//     PlcTask Inputs/GVL_iXlinker.Device_2_EtherCAT.Term_9_EK1100.Term_34_EL3403.PM_Inputs_Channel_1.TxPDO_Toggle <-> PM Inputs Channel 1/TxPDO Toggle
//     PlcTask Inputs/GVL_iXlinker.Device_2_EtherCAT.Term_9_EK1100.Term_34_EL3403.PM_Inputs_Channel_2.TxPDO_Toggle <-> PM Inputs Channel 2/TxPDO Toggle
//     PlcTask Inputs/GVL_iXlinker.Device_2_EtherCAT.Term_9_EK1100.Term_34_EL3403.PM_Inputs_Channel_3.TxPDO_Toggle <-> PM Inputs Channel 3/TxPDO Toggle
//     PlcTask Inputs/GVL_iXlinker.Device_2_EtherCAT.Term_9_EK1100.Term_34_EL3403.PM_Inputs_Channel_1.Variant_value <-> PM Inputs Channel 1/Variant value
//     PlcTask Inputs/GVL_iXlinker.Device_2_EtherCAT.Term_9_EK1100.Term_34_EL3403.PM_Inputs_Channel_2.Variant_value <-> PM Inputs Channel 2/Variant value
//     PlcTask Inputs/GVL_iXlinker.Device_2_EtherCAT.Term_9_EK1100.Term_34_EL3403.PM_Inputs_Channel_3.Variant_value <-> PM Inputs Channel 3/Variant value
//     PlcTask Inputs/GVL_iXlinker.Device_2_EtherCAT.Term_9_EK1100.Term_34_EL3403.PM_Inputs_Channel_1.Voltage <-> PM Inputs Channel 1/Voltage
//     PlcTask Inputs/GVL_iXlinker.Device_2_EtherCAT.Term_9_EK1100.Term_34_EL3403.PM_Inputs_Channel_2.Voltage <-> PM Inputs Channel 2/Voltage
//     PlcTask Inputs/GVL_iXlinker.Device_2_EtherCAT.Term_9_EK1100.Term_34_EL3403.PM_Inputs_Channel_3.Voltage <-> PM Inputs Channel 3/Voltage
//     PlcTask Inputs/GVL_iXlinker.Device_2_EtherCAT.Term_9_EK1100.Term_34_EL3403.PM_Status_data.Missing_zero_crossing_A <-> PM Status data/Missing zero crossing A
//     PlcTask Inputs/GVL_iXlinker.Device_2_EtherCAT.Term_9_EK1100.Term_34_EL3403.PM_Status_data.Missing_zero_crossing_B <-> PM Status data/Missing zero crossing B
//     PlcTask Inputs/GVL_iXlinker.Device_2_EtherCAT.Term_9_EK1100.Term_34_EL3403.PM_Status_data.Missing_zero_crossing_C <-> PM Status data/Missing zero crossing C
//     PlcTask Inputs/GVL_iXlinker.Device_2_EtherCAT.Term_9_EK1100.Term_34_EL3403.PM_Status_data.Phase_sequence_error <-> PM Status data/Phase sequence error
//     PlcTask Inputs/GVL_iXlinker.Device_2_EtherCAT.Term_9_EK1100.Term_34_EL3403.WcState.InputToggle <-> WcState/InputToggle
//     PlcTask Inputs/GVL_iXlinker.Device_2_EtherCAT.Term_9_EK1100.Term_34_EL3403.WcState.WcState <-> WcState/WcState
//     PlcTask Outputs/GVL_iXlinker.Device_2_EtherCAT.Term_9_EK1100.Term_34_EL3403.PM_Outputs_Channel_1.Index <-> PM Outputs Channel 1/Index
//     PlcTask Outputs/GVL_iXlinker.Device_2_EtherCAT.Term_9_EK1100.Term_34_EL3403.PM_Outputs_Channel_2.Index <-> PM Outputs Channel 2/Index
//     PlcTask Outputs/GVL_iXlinker.Device_2_EtherCAT.Term_9_EK1100.Term_34_EL3403.PM_Outputs_Channel_3.Index <-> PM Outputs Channel 3/Index
//   TcoIoTests/TcoIoTests Instance <-> Device 2 (EtherCAT)/Term 9 (EK1100)/Term 35 (EL6001)
//     PlcTask Inputs/GVL_iXlinker.Device_2_EtherCAT.Term_9_EK1100.Term_35_EL6001.COM_Inputs.Data_In[{0..21}] <-> COM Inputs/Data In {0..21}  (22 links)
//     PlcTask Inputs/GVL_iXlinker.Device_2_EtherCAT.Term_9_EK1100.Term_35_EL6001.COM_Inputs.Status/Buffer_full <-> COM Inputs/Status/Buffer full
//     PlcTask Inputs/GVL_iXlinker.Device_2_EtherCAT.Term_9_EK1100.Term_35_EL6001.COM_Inputs.Status/Framing_error <-> COM Inputs/Status/Framing error
//     PlcTask Inputs/GVL_iXlinker.Device_2_EtherCAT.Term_9_EK1100.Term_35_EL6001.COM_Inputs.Status/Init_accepted <-> COM Inputs/Status/Init accepted
//     PlcTask Inputs/GVL_iXlinker.Device_2_EtherCAT.Term_9_EK1100.Term_35_EL6001.COM_Inputs.Status/Input_length <-> COM Inputs/Status/Input length
//     PlcTask Inputs/GVL_iXlinker.Device_2_EtherCAT.Term_9_EK1100.Term_35_EL6001.COM_Inputs.Status/Overrun_error <-> COM Inputs/Status/Overrun error
//     PlcTask Inputs/GVL_iXlinker.Device_2_EtherCAT.Term_9_EK1100.Term_35_EL6001.COM_Inputs.Status/Parity_error <-> COM Inputs/Status/Parity error
//     PlcTask Inputs/GVL_iXlinker.Device_2_EtherCAT.Term_9_EK1100.Term_35_EL6001.COM_Inputs.Status/Receive_request <-> COM Inputs/Status/Receive request
//     PlcTask Inputs/GVL_iXlinker.Device_2_EtherCAT.Term_9_EK1100.Term_35_EL6001.COM_Inputs.Status/Transmit_accepted <-> COM Inputs/Status/Transmit accepted
//     PlcTask Inputs/GVL_iXlinker.Device_2_EtherCAT.Term_9_EK1100.Term_35_EL6001.InfoData.AdsAddr <-> InfoData/AdsAddr
//     PlcTask Inputs/GVL_iXlinker.Device_2_EtherCAT.Term_9_EK1100.Term_35_EL6001.InfoData.State <-> InfoData/State
//     PlcTask Inputs/GVL_iXlinker.Device_2_EtherCAT.Term_9_EK1100.Term_35_EL6001.WcState.InputToggle <-> WcState/InputToggle
//     PlcTask Inputs/GVL_iXlinker.Device_2_EtherCAT.Term_9_EK1100.Term_35_EL6001.WcState.WcState <-> WcState/WcState
//     PlcTask Outputs/GVL_iXlinker.Device_2_EtherCAT.Term_9_EK1100.Term_35_EL6001.COM_Outputs.Ctrl/Init_request <-> COM Outputs/Ctrl/Init request
//     PlcTask Outputs/GVL_iXlinker.Device_2_EtherCAT.Term_9_EK1100.Term_35_EL6001.COM_Outputs.Ctrl/Output_length <-> COM Outputs/Ctrl/Output length
//     PlcTask Outputs/GVL_iXlinker.Device_2_EtherCAT.Term_9_EK1100.Term_35_EL6001.COM_Outputs.Ctrl/Receive_accepted <-> COM Outputs/Ctrl/Receive accepted
//     PlcTask Outputs/GVL_iXlinker.Device_2_EtherCAT.Term_9_EK1100.Term_35_EL6001.COM_Outputs.Ctrl/Send_continues <-> COM Outputs/Ctrl/Send continues
//     PlcTask Outputs/GVL_iXlinker.Device_2_EtherCAT.Term_9_EK1100.Term_35_EL6001.COM_Outputs.Ctrl/Transmit_request <-> COM Outputs/Ctrl/Transmit request
//     PlcTask Outputs/GVL_iXlinker.Device_2_EtherCAT.Term_9_EK1100.Term_35_EL6001.COM_Outputs.Data_Out[{0..21}] <-> COM Outputs/Data Out {0..21}  (22 links)
//   TcoIoTests/TcoIoTests Instance <-> Device 2 (EtherCAT)/Term 9 (EK1100)/Term 36 (EL3024)
//     PlcTask Inputs/GVL_iXlinker.Device_2_EtherCAT.Term_9_EK1100.Term_36_EL3024.AI_Standard_Channel_{1..4}.Status/Error <-> AI Standard Channel {1..4}/Status/Error  (4 links)
//     PlcTask Inputs/GVL_iXlinker.Device_2_EtherCAT.Term_9_EK1100.Term_36_EL3024.AI_Standard_Channel_1.Status/Limit_1 <-> AI Standard Channel 1/Status/Limit 1
//     PlcTask Inputs/GVL_iXlinker.Device_2_EtherCAT.Term_9_EK1100.Term_36_EL3024.AI_Standard_Channel_1.Status/Limit_2 <-> AI Standard Channel 1/Status/Limit 2
//     PlcTask Inputs/GVL_iXlinker.Device_2_EtherCAT.Term_9_EK1100.Term_36_EL3024.AI_Standard_Channel_2.Status/Limit_1 <-> AI Standard Channel 2/Status/Limit 1
//     PlcTask Inputs/GVL_iXlinker.Device_2_EtherCAT.Term_9_EK1100.Term_36_EL3024.AI_Standard_Channel_2.Status/Limit_2 <-> AI Standard Channel 2/Status/Limit 2
//     PlcTask Inputs/GVL_iXlinker.Device_2_EtherCAT.Term_9_EK1100.Term_36_EL3024.AI_Standard_Channel_3.Status/Limit_1 <-> AI Standard Channel 3/Status/Limit 1
//     PlcTask Inputs/GVL_iXlinker.Device_2_EtherCAT.Term_9_EK1100.Term_36_EL3024.AI_Standard_Channel_3.Status/Limit_2 <-> AI Standard Channel 3/Status/Limit 2
//     PlcTask Inputs/GVL_iXlinker.Device_2_EtherCAT.Term_9_EK1100.Term_36_EL3024.AI_Standard_Channel_4.Status/Limit_1 <-> AI Standard Channel 4/Status/Limit 1
//     PlcTask Inputs/GVL_iXlinker.Device_2_EtherCAT.Term_9_EK1100.Term_36_EL3024.AI_Standard_Channel_4.Status/Limit_2 <-> AI Standard Channel 4/Status/Limit 2
//     PlcTask Inputs/GVL_iXlinker.Device_2_EtherCAT.Term_9_EK1100.Term_36_EL3024.AI_Standard_Channel_{1..4}.Status/Overrange <-> AI Standard Channel {1..4}/Status/Overrange  (4 links)
//     PlcTask Inputs/GVL_iXlinker.Device_2_EtherCAT.Term_9_EK1100.Term_36_EL3024.AI_Standard_Channel_{1..4}.Status/TxPDO_State <-> AI Standard Channel {1..4}/Status/TxPDO State  (4 links)
//     PlcTask Inputs/GVL_iXlinker.Device_2_EtherCAT.Term_9_EK1100.Term_36_EL3024.AI_Standard_Channel_{1..4}.Status/TxPDO_Toggle <-> AI Standard Channel {1..4}/Status/TxPDO Toggle  (4 links)
//     PlcTask Inputs/GVL_iXlinker.Device_2_EtherCAT.Term_9_EK1100.Term_36_EL3024.AI_Standard_Channel_{1..4}.Status/Underrange <-> AI Standard Channel {1..4}/Status/Underrange  (4 links)
//     PlcTask Inputs/GVL_iXlinker.Device_2_EtherCAT.Term_9_EK1100.Term_36_EL3024.AI_Standard_Channel_{1..4}.Value <-> AI Standard Channel {1..4}/Value  (4 links)
//     PlcTask Inputs/GVL_iXlinker.Device_2_EtherCAT.Term_9_EK1100.Term_36_EL3024.InfoData.AdsAddr <-> InfoData/AdsAddr
//     PlcTask Inputs/GVL_iXlinker.Device_2_EtherCAT.Term_9_EK1100.Term_36_EL3024.InfoData.State <-> InfoData/State
//     PlcTask Inputs/GVL_iXlinker.Device_2_EtherCAT.Term_9_EK1100.Term_36_EL3024.WcState.InputToggle <-> WcState/InputToggle
//     PlcTask Inputs/GVL_iXlinker.Device_2_EtherCAT.Term_9_EK1100.Term_36_EL3024.WcState.WcState <-> WcState/WcState
//   TcoIoTests/TcoIoTests Instance <-> Device 3 (EtherCAT)
//     PlcTask Inputs/GVL_iXlinker.Device_3_EtherCAT.InfoData.AmsNetId <-> InfoData/AmsNetId
//     PlcTask Inputs/GVL_iXlinker.Device_3_EtherCAT.InfoData.CfgSlaveCount <-> InfoData/CfgSlaveCount
//     PlcTask Inputs/GVL_iXlinker.Device_3_EtherCAT.InfoData.ChangeCount <-> InfoData/ChangeCount
//     PlcTask Inputs/GVL_iXlinker.Device_3_EtherCAT.InfoData.DevId <-> InfoData/DevId
//     PlcTask Inputs/GVL_iXlinker.Device_3_EtherCAT.Inputs.DevState <-> Inputs/DevState
//     PlcTask Inputs/GVL_iXlinker.Device_3_EtherCAT.Inputs.Frm0InputToggle <-> Inputs/Frm0InputToggle
//     PlcTask Inputs/GVL_iXlinker.Device_3_EtherCAT.Inputs.Frm0State <-> Inputs/Frm0State
//     PlcTask Inputs/GVL_iXlinker.Device_3_EtherCAT.Inputs.Frm0WcState <-> Inputs/Frm0WcState
//     PlcTask Inputs/GVL_iXlinker.Device_3_EtherCAT.Inputs.SlaveCount <-> Inputs/SlaveCount
//     PlcTask Outputs/GVL_iXlinker.Device_3_EtherCAT.Outputs.DevCtrl <-> Outputs/DevCtrl
//     PlcTask Outputs/GVL_iXlinker.Device_3_EtherCAT.Outputs.Frm0Ctrl <-> Outputs/Frm0Ctrl
//     PlcTask Outputs/GVL_iXlinker.Device_3_EtherCAT.Outputs.Frm0WcCtrl <-> Outputs/Frm0WcCtrl
//   TcoIoTests/TcoIoTests Instance <-> Device 3 (EtherCAT)/Term 146 (EK1100)
//     PlcTask Inputs/GVL_iXlinker.Device_3_EtherCAT.Term_146_EK1100.InfoData.State <-> InfoData/State
//   TcoIoTests/TcoIoTests Instance <-> Device 3 (EtherCAT)/Term 146 (EK1100)/Term 147 (EK1122)
//     PlcTask Inputs/GVL_iXlinker.Device_3_EtherCAT.Term_146_EK1100.Term_147_EK1122.InfoData.State <-> InfoData/State
//   TcoIoTests/TcoIoTests Instance <-> Device 3 (EtherCAT)/Term 146 (EK1100)/Term 147 (EK1122)/Term 153 (EK1100)
//     PlcTask Inputs/GVL_iXlinker.Device_3_EtherCAT.Term_146_EK1100.Term_147_EK1122.Term_153_EK1100.InfoData.State <-> InfoData/State
//   TcoIoTests/TcoIoTests Instance <-> Device 3 (EtherCAT)/Term 146 (EK1100)/Term 147 (EK1122)/Term 153 (EK1100)/Term 154 (EK1122)
//     PlcTask Inputs/GVL_iXlinker.Device_3_EtherCAT.Term_146_EK1100.Term_147_EK1122.Term_153_EK1100.Term_154_EK1122.InfoData.State <-> InfoData/State
//   TcoIoTests/TcoIoTests Instance <-> Device 3 (EtherCAT)/Term 146 (EK1100)/Term 147 (EK1122)/Term 153 (EK1100)/Term 154 (EK1122)/Term 157 (EK1100)
//     PlcTask Inputs/GVL_iXlinker.Device_3_EtherCAT.Term_146_EK1100.Term_147_EK1122.Term_153_EK1100.Term_154_EK1122.Term_157_EK1100.InfoData.State <-> InfoData/State
//   TcoIoTests/TcoIoTests Instance <-> Device 3 (EtherCAT)/Term 146 (EK1100)/Term 147 (EK1122)/Term 153 (EK1100)/Term 154 (EK1122)/Term 157 (EK1100)/Term 159 (EL1809)
//     PlcTask Inputs/GVL_iXlinker.Device_3_EtherCAT.Term_146_EK1100.Term_147_EK1122.Term_153_EK1100.Term_154_EK1122.Term_157_EK1100.Term_159_EL1809.Channel_{1..16}.Input <-> Channel {1..16}/Input  (16 links)
//     PlcTask Inputs/GVL_iXlinker.Device_3_EtherCAT.Term_146_EK1100.Term_147_EK1122.Term_153_EK1100.Term_154_EK1122.Term_157_EK1100.Term_159_EL1809.InfoData.State <-> InfoData/State
//     PlcTask Inputs/GVL_iXlinker.Device_3_EtherCAT.Term_146_EK1100.Term_147_EK1122.Term_153_EK1100.Term_154_EK1122.Term_157_EK1100.Term_159_EL1809.WcState.InputToggle <-> WcState/InputToggle
//     PlcTask Inputs/GVL_iXlinker.Device_3_EtherCAT.Term_146_EK1100.Term_147_EK1122.Term_153_EK1100.Term_154_EK1122.Term_157_EK1100.Term_159_EL1809.WcState.WcState <-> WcState/WcState
//   TcoIoTests/TcoIoTests Instance <-> Device 3 (EtherCAT)/Term 146 (EK1100)/Term 147 (EK1122)/Term 153 (EK1100)/Term 154 (EK1122)/Term 158 (EK1100)
//     PlcTask Inputs/GVL_iXlinker.Device_3_EtherCAT.Term_146_EK1100.Term_147_EK1122.Term_153_EK1100.Term_154_EK1122.Term_158_EK1100.InfoData.State <-> InfoData/State
//   TcoIoTests/TcoIoTests Instance <-> Device 3 (EtherCAT)/Term 146 (EK1100)/Term 147 (EK1122)/Term 153 (EK1100)/Term 154 (EK1122)/Term 158 (EK1100)/Term 160 (EL1809)
//     PlcTask Inputs/GVL_iXlinker.Device_3_EtherCAT.Term_146_EK1100.Term_147_EK1122.Term_153_EK1100.Term_154_EK1122.Term_158_EK1100.Term_160_EL1809.Channel_{1..16}.Input <-> Channel {1..16}/Input  (16 links)
//     PlcTask Inputs/GVL_iXlinker.Device_3_EtherCAT.Term_146_EK1100.Term_147_EK1122.Term_153_EK1100.Term_154_EK1122.Term_158_EK1100.Term_160_EL1809.InfoData.State <-> InfoData/State
//     PlcTask Inputs/GVL_iXlinker.Device_3_EtherCAT.Term_146_EK1100.Term_147_EK1122.Term_153_EK1100.Term_154_EK1122.Term_158_EK1100.Term_160_EL1809.WcState.InputToggle <-> WcState/InputToggle
//     PlcTask Inputs/GVL_iXlinker.Device_3_EtherCAT.Term_146_EK1100.Term_147_EK1122.Term_153_EK1100.Term_154_EK1122.Term_158_EK1100.Term_160_EL1809.WcState.WcState <-> WcState/WcState
//   TcoIoTests/TcoIoTests Instance <-> Device 3 (EtherCAT)/Term 146 (EK1100)/Term 147 (EK1122)/Term 153 (EK1100)/Term 155 (EL2008)
//     PlcTask Inputs/GVL_iXlinker.Device_3_EtherCAT.Term_146_EK1100.Term_147_EK1122.Term_153_EK1100.Term_155_EL2008.InfoData.State <-> InfoData/State
//     PlcTask Inputs/GVL_iXlinker.Device_3_EtherCAT.Term_146_EK1100.Term_147_EK1122.Term_153_EK1100.Term_155_EL2008.WcState.WcState <-> WcState/WcState
//     PlcTask Outputs/GVL_iXlinker.Device_3_EtherCAT.Term_146_EK1100.Term_147_EK1122.Term_153_EK1100.Term_155_EL2008.Channel_{1..8}.Output <-> Channel {1..8}/Output  (8 links)
//   TcoIoTests/TcoIoTests Instance <-> Device 3 (EtherCAT)/Term 146 (EK1100)/Term 147 (EK1122)/Term 153 (EK1100)/Term 156 (EL2008)
//     PlcTask Inputs/GVL_iXlinker.Device_3_EtherCAT.Term_146_EK1100.Term_147_EK1122.Term_153_EK1100.Term_156_EL2008.InfoData.State <-> InfoData/State
//     PlcTask Inputs/GVL_iXlinker.Device_3_EtherCAT.Term_146_EK1100.Term_147_EK1122.Term_153_EK1100.Term_156_EL2008.WcState.WcState <-> WcState/WcState
//     PlcTask Outputs/GVL_iXlinker.Device_3_EtherCAT.Term_146_EK1100.Term_147_EK1122.Term_153_EK1100.Term_156_EL2008.Channel_{1..8}.Output <-> Channel {1..8}/Output  (8 links)
//   TcoIoTests/TcoIoTests Instance <-> Device 3 (EtherCAT)/Term 146 (EK1100)/Term 147 (EK1122)/Term 178 (EK1100)
//     PlcTask Inputs/GVL_iXlinker.Device_3_EtherCAT.Term_146_EK1100.Term_147_EK1122.Term_178_EK1100.InfoData.State <-> InfoData/State
//   TcoIoTests/TcoIoTests Instance <-> Device 3 (EtherCAT)/Term 146 (EK1100)/Term 147 (EK1122)/Term 178 (EK1100)/Term 179 (EK1122)
//     PlcTask Inputs/GVL_iXlinker.Device_3_EtherCAT.Term_146_EK1100.Term_147_EK1122.Term_178_EK1100.Term_179_EK1122.InfoData.State <-> InfoData/State
//   TcoIoTests/TcoIoTests Instance <-> Device 3 (EtherCAT)/Term 146 (EK1100)/Term 147 (EK1122)/Term 178 (EK1100)/Term 179 (EK1122)/Term 180 (EK1100)
//     PlcTask Inputs/GVL_iXlinker.Device_3_EtherCAT.Term_146_EK1100.Term_147_EK1122.Term_178_EK1100.Term_179_EK1122.Term_180_EK1100.InfoData.State <-> InfoData/State
//   TcoIoTests/TcoIoTests Instance <-> Device 3 (EtherCAT)/Term 146 (EK1100)/Term 147 (EK1122)/Term 178 (EK1100)/Term 179 (EK1122)/Term 180 (EK1100)/Term 181 (EL1809)
//     PlcTask Inputs/GVL_iXlinker.Device_3_EtherCAT.Term_146_EK1100.Term_147_EK1122.Term_178_EK1100.Term_179_EK1122.Term_180_EK1100.Term_181_EL1809.Channel_{1..16}.Input <-> Channel {1..16}/Input  (16 links)
//     PlcTask Inputs/GVL_iXlinker.Device_3_EtherCAT.Term_146_EK1100.Term_147_EK1122.Term_178_EK1100.Term_179_EK1122.Term_180_EK1100.Term_181_EL1809.InfoData.State <-> InfoData/State
//     PlcTask Inputs/GVL_iXlinker.Device_3_EtherCAT.Term_146_EK1100.Term_147_EK1122.Term_178_EK1100.Term_179_EK1122.Term_180_EK1100.Term_181_EL1809.WcState.InputToggle <-> WcState/InputToggle
//     PlcTask Inputs/GVL_iXlinker.Device_3_EtherCAT.Term_146_EK1100.Term_147_EK1122.Term_178_EK1100.Term_179_EK1122.Term_180_EK1100.Term_181_EL1809.WcState.WcState <-> WcState/WcState
//   TcoIoTests/TcoIoTests Instance <-> Device 3 (EtherCAT)/Term 146 (EK1100)/Term 147 (EK1122)/Term 178 (EK1100)/Term 179 (EK1122)/Term 182 (EK1100)
//     PlcTask Inputs/GVL_iXlinker.Device_3_EtherCAT.Term_146_EK1100.Term_147_EK1122.Term_178_EK1100.Term_179_EK1122.Term_182_EK1100.InfoData.State <-> InfoData/State
//   TcoIoTests/TcoIoTests Instance <-> Device 3 (EtherCAT)/Term 146 (EK1100)/Term 147 (EK1122)/Term 178 (EK1100)/Term 179 (EK1122)/Term 182 (EK1100)/Term 183 (EL1809)
//     PlcTask Inputs/GVL_iXlinker.Device_3_EtherCAT.Term_146_EK1100.Term_147_EK1122.Term_178_EK1100.Term_179_EK1122.Term_182_EK1100.Term_183_EL1809.Channel_{1..16}.Input <-> Channel {1..16}/Input  (16 links)
//     PlcTask Inputs/GVL_iXlinker.Device_3_EtherCAT.Term_146_EK1100.Term_147_EK1122.Term_178_EK1100.Term_179_EK1122.Term_182_EK1100.Term_183_EL1809.InfoData.State <-> InfoData/State
//     PlcTask Inputs/GVL_iXlinker.Device_3_EtherCAT.Term_146_EK1100.Term_147_EK1122.Term_178_EK1100.Term_179_EK1122.Term_182_EK1100.Term_183_EL1809.WcState.InputToggle <-> WcState/InputToggle
//     PlcTask Inputs/GVL_iXlinker.Device_3_EtherCAT.Term_146_EK1100.Term_147_EK1122.Term_178_EK1100.Term_179_EK1122.Term_182_EK1100.Term_183_EL1809.WcState.WcState <-> WcState/WcState
//   TcoIoTests/TcoIoTests Instance <-> Device 3 (EtherCAT)/Term 146 (EK1100)/Term 147 (EK1122)/Term 178 (EK1100)/Term 184 (EL2008)
//     PlcTask Inputs/GVL_iXlinker.Device_3_EtherCAT.Term_146_EK1100.Term_147_EK1122.Term_178_EK1100.Term_184_EL2008.InfoData.State <-> InfoData/State
//     PlcTask Inputs/GVL_iXlinker.Device_3_EtherCAT.Term_146_EK1100.Term_147_EK1122.Term_178_EK1100.Term_184_EL2008.WcState.WcState <-> WcState/WcState
//     PlcTask Outputs/GVL_iXlinker.Device_3_EtherCAT.Term_146_EK1100.Term_147_EK1122.Term_178_EK1100.Term_184_EL2008.Channel_{1..8}.Output <-> Channel {1..8}/Output  (8 links)
//   TcoIoTests/TcoIoTests Instance <-> Device 3 (EtherCAT)/Term 146 (EK1100)/Term 147 (EK1122)/Term 178 (EK1100)/Term 185 (EL2008)
//     PlcTask Inputs/GVL_iXlinker.Device_3_EtherCAT.Term_146_EK1100.Term_147_EK1122.Term_178_EK1100.Term_185_EL2008.InfoData.State <-> InfoData/State
//     PlcTask Inputs/GVL_iXlinker.Device_3_EtherCAT.Term_146_EK1100.Term_147_EK1122.Term_178_EK1100.Term_185_EL2008.WcState.WcState <-> WcState/WcState
//     PlcTask Outputs/GVL_iXlinker.Device_3_EtherCAT.Term_146_EK1100.Term_147_EK1122.Term_178_EK1100.Term_185_EL2008.Channel_{1..8}.Output <-> Channel {1..8}/Output  (8 links)
//   TcoIoTests/TcoIoTests Instance <-> Device 3 (EtherCAT)/Term 146 (EK1100)/Term 148 (EL1809)
//     PlcTask Inputs/GVL_iXlinker.Device_3_EtherCAT.Term_146_EK1100.Term_148_EL1809.Channel_{1..16}.Input <-> Channel {1..16}/Input  (16 links)
//     PlcTask Inputs/GVL_iXlinker.Device_3_EtherCAT.Term_146_EK1100.Term_148_EL1809.InfoData.State <-> InfoData/State
//     PlcTask Inputs/GVL_iXlinker.Device_3_EtherCAT.Term_146_EK1100.Term_148_EL1809.WcState.InputToggle <-> WcState/InputToggle
//     PlcTask Inputs/GVL_iXlinker.Device_3_EtherCAT.Term_146_EK1100.Term_148_EL1809.WcState.WcState <-> WcState/WcState
//   TcoIoTests/TcoIoTests Instance <-> Device 3 (EtherCAT)/Term 146 (EK1100)/Term 149 (EL1809)
//     PlcTask Inputs/GVL_iXlinker.Device_3_EtherCAT.Term_146_EK1100.Term_149_EL1809.Channel_{1..16}.Input <-> Channel {1..16}/Input  (16 links)
//     PlcTask Inputs/GVL_iXlinker.Device_3_EtherCAT.Term_146_EK1100.Term_149_EL1809.InfoData.State <-> InfoData/State
//     PlcTask Inputs/GVL_iXlinker.Device_3_EtherCAT.Term_146_EK1100.Term_149_EL1809.WcState.InputToggle <-> WcState/InputToggle
//     PlcTask Inputs/GVL_iXlinker.Device_3_EtherCAT.Term_146_EK1100.Term_149_EL1809.WcState.WcState <-> WcState/WcState
//   TcoIoTests/TcoIoTests Instance <-> Device 3 (EtherCAT)/Term 146 (EK1100)/Term 150 (EL1809)
//     PlcTask Inputs/GVL_iXlinker.Device_3_EtherCAT.Term_146_EK1100.Term_150_EL1809.Channel_{1..16}.Input <-> Channel {1..16}/Input  (16 links)
//     PlcTask Inputs/GVL_iXlinker.Device_3_EtherCAT.Term_146_EK1100.Term_150_EL1809.InfoData.State <-> InfoData/State
//     PlcTask Inputs/GVL_iXlinker.Device_3_EtherCAT.Term_146_EK1100.Term_150_EL1809.WcState.InputToggle <-> WcState/InputToggle
//     PlcTask Inputs/GVL_iXlinker.Device_3_EtherCAT.Term_146_EK1100.Term_150_EL1809.WcState.WcState <-> WcState/WcState
//   TcoIoTests/TcoIoTests Instance <-> Device 3 (EtherCAT)/Term 146 (EK1100)/Term 151 (EL1809)
//     PlcTask Inputs/GVL_iXlinker.Device_3_EtherCAT.Term_146_EK1100.Term_151_EL1809.Channel_{1..16}.Input <-> Channel {1..16}/Input  (16 links)
//     PlcTask Inputs/GVL_iXlinker.Device_3_EtherCAT.Term_146_EK1100.Term_151_EL1809.InfoData.State <-> InfoData/State
//     PlcTask Inputs/GVL_iXlinker.Device_3_EtherCAT.Term_146_EK1100.Term_151_EL1809.WcState.InputToggle <-> WcState/InputToggle
//     PlcTask Inputs/GVL_iXlinker.Device_3_EtherCAT.Term_146_EK1100.Term_151_EL1809.WcState.WcState <-> WcState/WcState
//   TcoIoTests/TcoIoTests Instance <-> Device 3 (EtherCAT)/Term 146 (EK1100)/Term 152 (EL1809)
//     PlcTask Inputs/GVL_iXlinker.Device_3_EtherCAT.Term_146_EK1100.Term_152_EL1809.Channel_{1..16}.Input <-> Channel {1..16}/Input  (16 links)
//     PlcTask Inputs/GVL_iXlinker.Device_3_EtherCAT.Term_146_EK1100.Term_152_EL1809.InfoData.State <-> InfoData/State
//     PlcTask Inputs/GVL_iXlinker.Device_3_EtherCAT.Term_146_EK1100.Term_152_EL1809.WcState.InputToggle <-> WcState/InputToggle
//     PlcTask Inputs/GVL_iXlinker.Device_3_EtherCAT.Term_146_EK1100.Term_152_EL1809.WcState.WcState <-> WcState/WcState
//   TcoIoTests/TcoIoTests Instance <-> Device 3 (EtherCAT)/Term 146 (EK1100)/Term 186 (EK1122)
//     PlcTask Inputs/GVL_iXlinker.Device_3_EtherCAT.Term_146_EK1100.Term_186_EK1122.InfoData.State <-> InfoData/State
//   TcoIoTests/TcoIoTests Instance <-> Device 3 (EtherCAT)/Term 146 (EK1100)/Term 186 (EK1122)/Term 187 (EK1100)
//     PlcTask Inputs/GVL_iXlinker.Device_3_EtherCAT.Term_146_EK1100.Term_186_EK1122.Term_187_EK1100.InfoData.State <-> InfoData/State
//   TcoIoTests/TcoIoTests Instance <-> Device 3 (EtherCAT)/Term 146 (EK1100)/Term 186 (EK1122)/Term 187 (EK1100)/Term 188 (EK1122)
//     PlcTask Inputs/GVL_iXlinker.Device_3_EtherCAT.Term_146_EK1100.Term_186_EK1122.Term_187_EK1100.Term_188_EK1122.InfoData.State <-> InfoData/State
//   TcoIoTests/TcoIoTests Instance <-> Device 3 (EtherCAT)/Term 146 (EK1100)/Term 186 (EK1122)/Term 187 (EK1100)/Term 188 (EK1122)/Term 189 (EK1100)
//     PlcTask Inputs/GVL_iXlinker.Device_3_EtherCAT.Term_146_EK1100.Term_186_EK1122.Term_187_EK1100.Term_188_EK1122.Term_189_EK1100.InfoData.State <-> InfoData/State
//   TcoIoTests/TcoIoTests Instance <-> Device 3 (EtherCAT)/Term 146 (EK1100)/Term 186 (EK1122)/Term 187 (EK1100)/Term 188 (EK1122)/Term 189 (EK1100)/Term 193 (EL1809)
//     PlcTask Inputs/GVL_iXlinker.Device_3_EtherCAT.Term_146_EK1100.Term_186_EK1122.Term_187_EK1100.Term_188_EK1122.Term_189_EK1100.Term_193_EL1809.Channel_{1..16}.Input <-> Channel {1..16}/Input  (16 links)
//     PlcTask Inputs/GVL_iXlinker.Device_3_EtherCAT.Term_146_EK1100.Term_186_EK1122.Term_187_EK1100.Term_188_EK1122.Term_189_EK1100.Term_193_EL1809.InfoData.State <-> InfoData/State
//     PlcTask Inputs/GVL_iXlinker.Device_3_EtherCAT.Term_146_EK1100.Term_186_EK1122.Term_187_EK1100.Term_188_EK1122.Term_189_EK1100.Term_193_EL1809.WcState.InputToggle <-> WcState/InputToggle
//     PlcTask Inputs/GVL_iXlinker.Device_3_EtherCAT.Term_146_EK1100.Term_186_EK1122.Term_187_EK1100.Term_188_EK1122.Term_189_EK1100.Term_193_EL1809.WcState.WcState <-> WcState/WcState
//   TcoIoTests/TcoIoTests Instance <-> Device 3 (EtherCAT)/Term 146 (EK1100)/Term 186 (EK1122)/Term 187 (EK1100)/Term 188 (EK1122)/Term 194 (EK1100)
//     PlcTask Inputs/GVL_iXlinker.Device_3_EtherCAT.Term_146_EK1100.Term_186_EK1122.Term_187_EK1100.Term_188_EK1122.Term_194_EK1100.InfoData.State <-> InfoData/State
//   TcoIoTests/TcoIoTests Instance <-> Device 3 (EtherCAT)/Term 146 (EK1100)/Term 186 (EK1122)/Term 187 (EK1100)/Term 188 (EK1122)/Term 194 (EK1100)/Term 200 (EL1809)
//     PlcTask Inputs/GVL_iXlinker.Device_3_EtherCAT.Term_146_EK1100.Term_186_EK1122.Term_187_EK1100.Term_188_EK1122.Term_194_EK1100.Term_200_EL1809.Channel_{1..16}.Input <-> Channel {1..16}/Input  (16 links)
//     PlcTask Inputs/GVL_iXlinker.Device_3_EtherCAT.Term_146_EK1100.Term_186_EK1122.Term_187_EK1100.Term_188_EK1122.Term_194_EK1100.Term_200_EL1809.InfoData.State <-> InfoData/State
//     PlcTask Inputs/GVL_iXlinker.Device_3_EtherCAT.Term_146_EK1100.Term_186_EK1122.Term_187_EK1100.Term_188_EK1122.Term_194_EK1100.Term_200_EL1809.WcState.InputToggle <-> WcState/InputToggle
//     PlcTask Inputs/GVL_iXlinker.Device_3_EtherCAT.Term_146_EK1100.Term_186_EK1122.Term_187_EK1100.Term_188_EK1122.Term_194_EK1100.Term_200_EL1809.WcState.WcState <-> WcState/WcState
//   TcoIoTests/TcoIoTests Instance <-> Device 3 (EtherCAT)/Term 146 (EK1100)/Term 186 (EK1122)/Term 187 (EK1100)/Term 204 (EL2008)
//     PlcTask Inputs/GVL_iXlinker.Device_3_EtherCAT.Term_146_EK1100.Term_186_EK1122.Term_187_EK1100.Term_204_EL2008.InfoData.State <-> InfoData/State
//     PlcTask Inputs/GVL_iXlinker.Device_3_EtherCAT.Term_146_EK1100.Term_186_EK1122.Term_187_EK1100.Term_204_EL2008.WcState.WcState <-> WcState/WcState
//     PlcTask Outputs/GVL_iXlinker.Device_3_EtherCAT.Term_146_EK1100.Term_186_EK1122.Term_187_EK1100.Term_204_EL2008.Channel_{1..8}.Output <-> Channel {1..8}/Output  (8 links)
//   TcoIoTests/TcoIoTests Instance <-> Device 3 (EtherCAT)/Term 146 (EK1100)/Term 186 (EK1122)/Term 187 (EK1100)/Term 205 (EL2008)
//     PlcTask Inputs/GVL_iXlinker.Device_3_EtherCAT.Term_146_EK1100.Term_186_EK1122.Term_187_EK1100.Term_205_EL2008.InfoData.State <-> InfoData/State
//     PlcTask Inputs/GVL_iXlinker.Device_3_EtherCAT.Term_146_EK1100.Term_186_EK1122.Term_187_EK1100.Term_205_EL2008.WcState.WcState <-> WcState/WcState
//     PlcTask Outputs/GVL_iXlinker.Device_3_EtherCAT.Term_146_EK1100.Term_186_EK1122.Term_187_EK1100.Term_205_EL2008.Channel_{1..8}.Output <-> Channel {1..8}/Output  (8 links)
//   TcoIoTests/TcoIoTests Instance <-> Device 3 (EtherCAT)/Term 146 (EK1100)/Term 186 (EK1122)/Term 207 (EK1100)
//     PlcTask Inputs/GVL_iXlinker.Device_3_EtherCAT.Term_146_EK1100.Term_186_EK1122.Term_207_EK1100.InfoData.State <-> InfoData/State
//   TcoIoTests/TcoIoTests Instance <-> Device 3 (EtherCAT)/Term 146 (EK1100)/Term 186 (EK1122)/Term 207 (EK1100)/Term 230 (EK1122)
//     PlcTask Inputs/GVL_iXlinker.Device_3_EtherCAT.Term_146_EK1100.Term_186_EK1122.Term_207_EK1100.Term_230_EK1122.InfoData.State <-> InfoData/State
//   TcoIoTests/TcoIoTests Instance <-> Device 3 (EtherCAT)/Term 146 (EK1100)/Term 186 (EK1122)/Term 207 (EK1100)/Term 230 (EK1122)/Term 231 (EK1100)
//     PlcTask Inputs/GVL_iXlinker.Device_3_EtherCAT.Term_146_EK1100.Term_186_EK1122.Term_207_EK1100.Term_230_EK1122.Term_231_EK1100.InfoData.State <-> InfoData/State
//   TcoIoTests/TcoIoTests Instance <-> Device 3 (EtherCAT)/Term 146 (EK1100)/Term 186 (EK1122)/Term 207 (EK1100)/Term 230 (EK1122)/Term 231 (EK1100)/Term 232 (EL1809)
//     PlcTask Inputs/GVL_iXlinker.Device_3_EtherCAT.Term_146_EK1100.Term_186_EK1122.Term_207_EK1100.Term_230_EK1122.Term_231_EK1100.Term_232_EL1809.Channel_{1..16}.Input <-> Channel {1..16}/Input  (16 links)
//     PlcTask Inputs/GVL_iXlinker.Device_3_EtherCAT.Term_146_EK1100.Term_186_EK1122.Term_207_EK1100.Term_230_EK1122.Term_231_EK1100.Term_232_EL1809.InfoData.State <-> InfoData/State
//     PlcTask Inputs/GVL_iXlinker.Device_3_EtherCAT.Term_146_EK1100.Term_186_EK1122.Term_207_EK1100.Term_230_EK1122.Term_231_EK1100.Term_232_EL1809.WcState.InputToggle <-> WcState/InputToggle
//     PlcTask Inputs/GVL_iXlinker.Device_3_EtherCAT.Term_146_EK1100.Term_186_EK1122.Term_207_EK1100.Term_230_EK1122.Term_231_EK1100.Term_232_EL1809.WcState.WcState <-> WcState/WcState
//   TcoIoTests/TcoIoTests Instance <-> Device 3 (EtherCAT)/Term 146 (EK1100)/Term 186 (EK1122)/Term 207 (EK1100)/Term 230 (EK1122)/Term 233 (EK1100)
//     PlcTask Inputs/GVL_iXlinker.Device_3_EtherCAT.Term_146_EK1100.Term_186_EK1122.Term_207_EK1100.Term_230_EK1122.Term_233_EK1100.InfoData.State <-> InfoData/State
//   TcoIoTests/TcoIoTests Instance <-> Device 3 (EtherCAT)/Term 146 (EK1100)/Term 186 (EK1122)/Term 207 (EK1100)/Term 230 (EK1122)/Term 233 (EK1100)/Term 234 (EL1809)
//     PlcTask Inputs/GVL_iXlinker.Device_3_EtherCAT.Term_146_EK1100.Term_186_EK1122.Term_207_EK1100.Term_230_EK1122.Term_233_EK1100.Term_234_EL1809.Channel_{1..16}.Input <-> Channel {1..16}/Input  (16 links)
//     PlcTask Inputs/GVL_iXlinker.Device_3_EtherCAT.Term_146_EK1100.Term_186_EK1122.Term_207_EK1100.Term_230_EK1122.Term_233_EK1100.Term_234_EL1809.InfoData.State <-> InfoData/State
//     PlcTask Inputs/GVL_iXlinker.Device_3_EtherCAT.Term_146_EK1100.Term_186_EK1122.Term_207_EK1100.Term_230_EK1122.Term_233_EK1100.Term_234_EL1809.WcState.InputToggle <-> WcState/InputToggle
//     PlcTask Inputs/GVL_iXlinker.Device_3_EtherCAT.Term_146_EK1100.Term_186_EK1122.Term_207_EK1100.Term_230_EK1122.Term_233_EK1100.Term_234_EL1809.WcState.WcState <-> WcState/WcState
//   TcoIoTests/TcoIoTests Instance <-> Device 3 (EtherCAT)/Term 146 (EK1100)/Term 186 (EK1122)/Term 207 (EK1100)/Term 235 (EL2008)
//     PlcTask Inputs/GVL_iXlinker.Device_3_EtherCAT.Term_146_EK1100.Term_186_EK1122.Term_207_EK1100.Term_235_EL2008.InfoData.State <-> InfoData/State
//     PlcTask Inputs/GVL_iXlinker.Device_3_EtherCAT.Term_146_EK1100.Term_186_EK1122.Term_207_EK1100.Term_235_EL2008.WcState.WcState <-> WcState/WcState
//     PlcTask Outputs/GVL_iXlinker.Device_3_EtherCAT.Term_146_EK1100.Term_186_EK1122.Term_207_EK1100.Term_235_EL2008.Channel_{1..8}.Output <-> Channel {1..8}/Output  (8 links)
//   TcoIoTests/TcoIoTests Instance <-> Device 3 (EtherCAT)/Term 146 (EK1100)/Term 186 (EK1122)/Term 207 (EK1100)/Term 236 (EL2008)
//     PlcTask Inputs/GVL_iXlinker.Device_3_EtherCAT.Term_146_EK1100.Term_186_EK1122.Term_207_EK1100.Term_236_EL2008.InfoData.State <-> InfoData/State
//     PlcTask Inputs/GVL_iXlinker.Device_3_EtherCAT.Term_146_EK1100.Term_186_EK1122.Term_207_EK1100.Term_236_EL2008.WcState.WcState <-> WcState/WcState
//     PlcTask Outputs/GVL_iXlinker.Device_3_EtherCAT.Term_146_EK1100.Term_186_EK1122.Term_207_EK1100.Term_236_EL2008.Channel_{1..8}.Output <-> Channel {1..8}/Output  (8 links)
//   TcoIoTests/TcoIoTests Instance <-> Device 3 (EtherCAT)/Term 146 (EK1100)/Term 288 (EK1122)
//     PlcTask Inputs/GVL_iXlinker.Device_3_EtherCAT.Term_146_EK1100.Term_288_EK1122.InfoData.State <-> InfoData/State
//   TcoIoTests/TcoIoTests Instance <-> Device 3 (EtherCAT)/Term 146 (EK1100)/Term 288 (EK1122)/Term 289 (EK1100)
//     PlcTask Inputs/GVL_iXlinker.Device_3_EtherCAT.Term_146_EK1100.Term_288_EK1122.Term_289_EK1100.InfoData.State <-> InfoData/State
//   TcoIoTests/TcoIoTests Instance <-> Device 3 (EtherCAT)/Term 146 (EK1100)/Term 288 (EK1122)/Term 289 (EK1100)/Term 237 (EK1122)
//     PlcTask Inputs/GVL_iXlinker.Device_3_EtherCAT.Term_146_EK1100.Term_288_EK1122.Term_289_EK1100.Term_237_EK1122.InfoData.State <-> InfoData/State
//   TcoIoTests/TcoIoTests Instance <-> Device 3 (EtherCAT)/Term 146 (EK1100)/Term 288 (EK1122)/Term 289 (EK1100)/Term 237 (EK1122)/Drive 238 (AX5101-0000-0214)
//     PlcTask Inputs/GVL_iXlinker.Device_3_EtherCAT.Term_146_EK1100.Term_288_EK1122.Term_289_EK1100.Term_237_EK1122.Drive_238_AX5101_0000_0214.AT_x.Drive_status_word <-> AT/Drive status word
//     PlcTask Inputs/GVL_iXlinker.Device_3_EtherCAT.Term_146_EK1100.Term_288_EK1122.Term_289_EK1100.Term_237_EK1122.Drive_238_AX5101_0000_0214.AT_x.Following_distance <-> AT/Following distance
//     PlcTask Inputs/GVL_iXlinker.Device_3_EtherCAT.Term_146_EK1100.Term_288_EK1122.Term_289_EK1100.Term_237_EK1122.Drive_238_AX5101_0000_0214.AT_x.Position_feedback_1_value <-> AT/Position feedback 1 value
//     PlcTask Inputs/GVL_iXlinker.Device_3_EtherCAT.Term_146_EK1100.Term_288_EK1122.Term_289_EK1100.Term_237_EK1122.Drive_238_AX5101_0000_0214.InfoData.AdsAddr <-> InfoData/AdsAddr
//     PlcTask Inputs/GVL_iXlinker.Device_3_EtherCAT.Term_146_EK1100.Term_288_EK1122.Term_289_EK1100.Term_237_EK1122.Drive_238_AX5101_0000_0214.InfoData.Chn0 <-> InfoData/Chn0
//     PlcTask Inputs/GVL_iXlinker.Device_3_EtherCAT.Term_146_EK1100.Term_288_EK1122.Term_289_EK1100.Term_237_EK1122.Drive_238_AX5101_0000_0214.InfoData.DcInputShift <-> InfoData/DcInputShift
//     PlcTask Inputs/GVL_iXlinker.Device_3_EtherCAT.Term_146_EK1100.Term_288_EK1122.Term_289_EK1100.Term_237_EK1122.Drive_238_AX5101_0000_0214.InfoData.DcOutputShift <-> InfoData/DcOutputShift
//     PlcTask Inputs/GVL_iXlinker.Device_3_EtherCAT.Term_146_EK1100.Term_288_EK1122.Term_289_EK1100.Term_237_EK1122.Drive_238_AX5101_0000_0214.InfoData.State <-> InfoData/State
//     PlcTask Inputs/GVL_iXlinker.Device_3_EtherCAT.Term_146_EK1100.Term_288_EK1122.Term_289_EK1100.Term_237_EK1122.Drive_238_AX5101_0000_0214.WcState.InputToggle <-> WcState/InputToggle
//     PlcTask Inputs/GVL_iXlinker.Device_3_EtherCAT.Term_146_EK1100.Term_288_EK1122.Term_289_EK1100.Term_237_EK1122.Drive_238_AX5101_0000_0214.WcState.WcState <-> WcState/WcState
//     PlcTask Outputs/GVL_iXlinker.Device_3_EtherCAT.Term_146_EK1100.Term_288_EK1122.Term_289_EK1100.Term_237_EK1122.Drive_238_AX5101_0000_0214.MDT.Master_control_word <-> MDT/Master control word
//     PlcTask Outputs/GVL_iXlinker.Device_3_EtherCAT.Term_146_EK1100.Term_288_EK1122.Term_289_EK1100.Term_237_EK1122.Drive_238_AX5101_0000_0214.MDT.Position_command_value <-> MDT/Position command value
//   TcoIoTests/TcoIoTests Instance <-> Device 3 (EtherCAT)/Term 146 (EK1100)/Term 288 (EK1122)/Term 289 (EK1100)/Term 293 (EL1809)
//     PlcTask Inputs/GVL_iXlinker.Device_3_EtherCAT.Term_146_EK1100.Term_288_EK1122.Term_289_EK1100.Term_293_EL1809.Channel_{1..16}.Input <-> Channel {1..16}/Input  (16 links)
//     PlcTask Inputs/GVL_iXlinker.Device_3_EtherCAT.Term_146_EK1100.Term_288_EK1122.Term_289_EK1100.Term_293_EL1809.InfoData.State <-> InfoData/State
//     PlcTask Inputs/GVL_iXlinker.Device_3_EtherCAT.Term_146_EK1100.Term_288_EK1122.Term_289_EK1100.Term_293_EL1809.WcState.InputToggle <-> WcState/InputToggle
//     PlcTask Inputs/GVL_iXlinker.Device_3_EtherCAT.Term_146_EK1100.Term_288_EK1122.Term_289_EK1100.Term_293_EL1809.WcState.WcState <-> WcState/WcState
//   TcoIoTests/TcoIoTests Instance <-> Device 3 (EtherCAT)/Term 146 (EK1100)/Term 288 (EK1122)/Term 294 (EK1100)
//     PlcTask Inputs/GVL_iXlinker.Device_3_EtherCAT.Term_146_EK1100.Term_288_EK1122.Term_294_EK1100.InfoData.State <-> InfoData/State
//   TcoIoTests/TcoIoTests Instance <-> Device 3 (EtherCAT)/Term 146 (EK1100)/Term 288 (EK1122)/Term 294 (EK1100)/Term 300 (EL1809)
//     PlcTask Inputs/GVL_iXlinker.Device_3_EtherCAT.Term_146_EK1100.Term_288_EK1122.Term_294_EK1100.Term_300_EL1809.Channel_{1..16}.Input <-> Channel {1..16}/Input  (16 links)
//     PlcTask Inputs/GVL_iXlinker.Device_3_EtherCAT.Term_146_EK1100.Term_288_EK1122.Term_294_EK1100.Term_300_EL1809.InfoData.State <-> InfoData/State
//     PlcTask Inputs/GVL_iXlinker.Device_3_EtherCAT.Term_146_EK1100.Term_288_EK1122.Term_294_EK1100.Term_300_EL1809.WcState.InputToggle <-> WcState/InputToggle
//     PlcTask Inputs/GVL_iXlinker.Device_3_EtherCAT.Term_146_EK1100.Term_288_EK1122.Term_294_EK1100.Term_300_EL1809.WcState.WcState <-> WcState/WcState
//   TcoIoTests/TcoIoTests Instance <-> Device 3 (EtherCAT)/Term 146 (EK1100)/Term 288 (EK1122)/Term 294 (EK1100)/Term 304 (EL2008)
//     PlcTask Inputs/GVL_iXlinker.Device_3_EtherCAT.Term_146_EK1100.Term_288_EK1122.Term_294_EK1100.Term_304_EL2008.InfoData.State <-> InfoData/State
//     PlcTask Inputs/GVL_iXlinker.Device_3_EtherCAT.Term_146_EK1100.Term_288_EK1122.Term_294_EK1100.Term_304_EL2008.WcState.WcState <-> WcState/WcState
//     PlcTask Outputs/GVL_iXlinker.Device_3_EtherCAT.Term_146_EK1100.Term_288_EK1122.Term_294_EK1100.Term_304_EL2008.Channel_{1..8}.Output <-> Channel {1..8}/Output  (8 links)
//   TcoIoTests/TcoIoTests Instance <-> Device 3 (EtherCAT)/Term 146 (EK1100)/Term 288 (EK1122)/Term 294 (EK1100)/Term 305 (EL2008)
//     PlcTask Inputs/GVL_iXlinker.Device_3_EtherCAT.Term_146_EK1100.Term_288_EK1122.Term_294_EK1100.Term_305_EL2008.InfoData.State <-> InfoData/State
//     PlcTask Inputs/GVL_iXlinker.Device_3_EtherCAT.Term_146_EK1100.Term_288_EK1122.Term_294_EK1100.Term_305_EL2008.WcState.WcState <-> WcState/WcState
//     PlcTask Outputs/GVL_iXlinker.Device_3_EtherCAT.Term_146_EK1100.Term_288_EK1122.Term_294_EK1100.Term_305_EL2008.Channel_{1..8}.Output <-> Channel {1..8}/Output  (8 links)
//   TcoIoTests/TcoIoTests Instance <-> Device 3 (EtherCAT)/Term 146 (EK1100)/Term 288 (EK1122)/Term 307 (EK1100)
//     PlcTask Inputs/GVL_iXlinker.Device_3_EtherCAT.Term_146_EK1100.Term_288_EK1122.Term_307_EK1100.InfoData.State <-> InfoData/State
//   TcoIoTests/TcoIoTests Instance <-> Device 3 (EtherCAT)/Term 146 (EK1100)/Term 288 (EK1122)/Term 307 (EK1100)/Term 330 (EK1122)
//     PlcTask Inputs/GVL_iXlinker.Device_3_EtherCAT.Term_146_EK1100.Term_288_EK1122.Term_307_EK1100.Term_330_EK1122.InfoData.State <-> InfoData/State
//   TcoIoTests/TcoIoTests Instance <-> Device 3 (EtherCAT)/Term 146 (EK1100)/Term 288 (EK1122)/Term 307 (EK1100)/Term 330 (EK1122)/Term 331 (EK1100)
//     PlcTask Inputs/GVL_iXlinker.Device_3_EtherCAT.Term_146_EK1100.Term_288_EK1122.Term_307_EK1100.Term_330_EK1122.Term_331_EK1100.InfoData.State <-> InfoData/State
//   TcoIoTests/TcoIoTests Instance <-> Device 3 (EtherCAT)/Term 146 (EK1100)/Term 288 (EK1122)/Term 307 (EK1100)/Term 330 (EK1122)/Term 331 (EK1100)/Term 332 (EL1809)
//     PlcTask Inputs/GVL_iXlinker.Device_3_EtherCAT.Term_146_EK1100.Term_288_EK1122.Term_307_EK1100.Term_330_EK1122.Term_331_EK1100.Term_332_EL1809.Channel_{1..16}.Input <-> Channel {1..16}/Input  (16 links)
//     PlcTask Inputs/GVL_iXlinker.Device_3_EtherCAT.Term_146_EK1100.Term_288_EK1122.Term_307_EK1100.Term_330_EK1122.Term_331_EK1100.Term_332_EL1809.InfoData.State <-> InfoData/State
//     PlcTask Inputs/GVL_iXlinker.Device_3_EtherCAT.Term_146_EK1100.Term_288_EK1122.Term_307_EK1100.Term_330_EK1122.Term_331_EK1100.Term_332_EL1809.WcState.InputToggle <-> WcState/InputToggle
//     PlcTask Inputs/GVL_iXlinker.Device_3_EtherCAT.Term_146_EK1100.Term_288_EK1122.Term_307_EK1100.Term_330_EK1122.Term_331_EK1100.Term_332_EL1809.WcState.WcState <-> WcState/WcState
//   TcoIoTests/TcoIoTests Instance <-> Device 3 (EtherCAT)/Term 146 (EK1100)/Term 288 (EK1122)/Term 307 (EK1100)/Term 330 (EK1122)/Term 333 (EK1100)
//     PlcTask Inputs/GVL_iXlinker.Device_3_EtherCAT.Term_146_EK1100.Term_288_EK1122.Term_307_EK1100.Term_330_EK1122.Term_333_EK1100.InfoData.State <-> InfoData/State
//   TcoIoTests/TcoIoTests Instance <-> Device 3 (EtherCAT)/Term 146 (EK1100)/Term 288 (EK1122)/Term 307 (EK1100)/Term 330 (EK1122)/Term 333 (EK1100)/Term 334 (EL1809)
//     PlcTask Inputs/GVL_iXlinker.Device_3_EtherCAT.Term_146_EK1100.Term_288_EK1122.Term_307_EK1100.Term_330_EK1122.Term_333_EK1100.Term_334_EL1809.Channel_{1..16}.Input <-> Channel {1..16}/Input  (16 links)
//     PlcTask Inputs/GVL_iXlinker.Device_3_EtherCAT.Term_146_EK1100.Term_288_EK1122.Term_307_EK1100.Term_330_EK1122.Term_333_EK1100.Term_334_EL1809.InfoData.State <-> InfoData/State
//     PlcTask Inputs/GVL_iXlinker.Device_3_EtherCAT.Term_146_EK1100.Term_288_EK1122.Term_307_EK1100.Term_330_EK1122.Term_333_EK1100.Term_334_EL1809.WcState.InputToggle <-> WcState/InputToggle
//     PlcTask Inputs/GVL_iXlinker.Device_3_EtherCAT.Term_146_EK1100.Term_288_EK1122.Term_307_EK1100.Term_330_EK1122.Term_333_EK1100.Term_334_EL1809.WcState.WcState <-> WcState/WcState
//   TcoIoTests/TcoIoTests Instance <-> Device 3 (EtherCAT)/Term 146 (EK1100)/Term 288 (EK1122)/Term 307 (EK1100)/Term 335 (EL2008)
//     PlcTask Inputs/GVL_iXlinker.Device_3_EtherCAT.Term_146_EK1100.Term_288_EK1122.Term_307_EK1100.Term_335_EL2008.InfoData.State <-> InfoData/State
//     PlcTask Inputs/GVL_iXlinker.Device_3_EtherCAT.Term_146_EK1100.Term_288_EK1122.Term_307_EK1100.Term_335_EL2008.WcState.WcState <-> WcState/WcState
//     PlcTask Outputs/GVL_iXlinker.Device_3_EtherCAT.Term_146_EK1100.Term_288_EK1122.Term_307_EK1100.Term_335_EL2008.Channel_{1..8}.Output <-> Channel {1..8}/Output  (8 links)
//   TcoIoTests/TcoIoTests Instance <-> Device 3 (EtherCAT)/Term 146 (EK1100)/Term 288 (EK1122)/Term 307 (EK1100)/Term 336 (EL2008)
//     PlcTask Inputs/GVL_iXlinker.Device_3_EtherCAT.Term_146_EK1100.Term_288_EK1122.Term_307_EK1100.Term_336_EL2008.InfoData.State <-> InfoData/State
//     PlcTask Inputs/GVL_iXlinker.Device_3_EtherCAT.Term_146_EK1100.Term_288_EK1122.Term_307_EK1100.Term_336_EL2008.WcState.WcState <-> WcState/WcState
//     PlcTask Outputs/GVL_iXlinker.Device_3_EtherCAT.Term_146_EK1100.Term_288_EK1122.Term_307_EK1100.Term_336_EL2008.Channel_{1..8}.Output <-> Channel {1..8}/Output  (8 links)

CONFIGURATION TcoIo
    RESOURCE PLC ON TwinCAT3
        TASK PlcTask(INTERVAL := T#15ms, PRIORITY := 12);
        PROGRAM MAIN WITH PlcTask : MAIN;
    END_RESOURCE
END_CONFIGURATION

// ---- Diagnostics/EtherCAT/MasterDevice/Base/EtcMasterBase_62654B43.TcDUT

TYPE EtcMasterBase_62654B43 :
STRUCT
END_STRUCT
END_TYPE

// ---- Diagnostics/EtherCAT/MasterDevice/Base/SyncUnitsBase_AD6C35CE.TcDUT

TYPE SyncUnitsBase_AD6C35CE :
STRUCT
END_STRUCT
END_TYPE

// ---- Diagnostics/EtherCAT/MasterDevice/Base/SyncUnitTaskBase_FCD3CBF3.TcDUT

TYPE SyncUnitTaskBase_FCD3CBF3 :
STRUCT
END_STRUCT
END_TYPE

// ---- Diagnostics/EtherCAT/MasterDevice/Base/SyncUnitTasksBase_7C8711EB.TcDUT

TYPE SyncUnitTasksBase_7C8711EB :
STRUCT
END_STRUCT
END_TYPE

// ---- Diagnostics/EtherCAT/MasterDevice/SyncUnit/InfoData_8649EEEB.TcDUT
{attribute 'GeneratedUsingTerminal: IODEVICETYPE_ETHERCATPROT'}
{attribute addProperty BoxType "IODEVICETYPE_ETHERCATPROT"}
{attribute addProperty Id "ObjectIdAT %I*DWORD4StateAT %I*UINT2SlaveCountAT %I*UINT2"}
{attribute addProperty CRC "2252992235"}
{attribute addProperty Size "8"}
TYPE InfoData_8649EEEB :
STRUCT
	{attribute addProperty Name "ObjectId"}
	ObjectId AT %I* : DWORD;
	{attribute addProperty Name "State"}
	State AT %I* : UINT;
	{attribute addProperty Name "SlaveCount"}
	SlaveCount AT %I* : UINT;
END_STRUCT
END_TYPE

// ---- Diagnostics/EtherCAT/MasterDevice/SyncUnit/SyncUnitState.TcDUT
TYPE SyncUnitState :
STRUCT
	{attribute addProperty Name "At least one slave in 'INIT' state"}	
    AtLeastOneSlaveInInitState : BOOL;
	{attribute addProperty Name "At least one slave in 'PREOP' state"}	
    AtLeastOneSlaveInPreopState : BOOL;
	{attribute addProperty Name "At least one slave in 'BOOT' state"}	
    AtLeastOneSlaveInBootState : BOOL;
	{attribute addProperty Name "At least one slave in 'SAFEOP' state"}	
    AtLeastOneSlaveInSafeOpState : BOOL;
	{attribute addProperty Name "At least one slave in 'OP' state"}	
    AtLeastOneSlaveInOpState : BOOL;
	{attribute addProperty Name "At least one slave signals error"}	
    AtLeastOneSlaveSignalsError : BOOL;
	{attribute addProperty Name "Invalid vendorId, productCode... read"}	
    InvalidVendoridOrProductcodeRead : BOOL;
	{attribute addProperty Name "Initialization error occurred"}	
    InitializationErrorOccurred : BOOL;
	{attribute addProperty Name "At least one slave disabled"}	
    AtLeastOneSlaveDisabled : BOOL;
	{attribute addProperty Name "At least one slave not present"}	
    AtLeastOneSlaveNotPresent : BOOL;
	{attribute addProperty Name "At least one slave signals link error"}	
    AtLeastOneSlaveSignalsLinkError : BOOL;
	{attribute addProperty Name "At least one slave signals missing link"}	
    AtLeastOneSlaveSignalsMissingLink : BOOL;
	{attribute addProperty Name "At least one slave signals unexpected link"}	
    AtLeastOneSlaveSignalsUnexpectedLink : BOOL;	
END_STRUCT
END_TYPE

// ---- Diagnostics/EtherCAT/MasterDevice/SyncUnit/SyncUnitTask_AB2F5079.TcDUT
{attribute 'GeneratedUsingTerminal: IODEVICETYPE_ETHERCATPROT'}
{attribute addProperty BoxType "IODEVICETYPE_ETHERCATPROT"}
{attribute addProperty Id "WcStateAT %I*WcState_0B2B16F91InfoDataAT %I*InfoData_8649EEEB8"}
{attribute addProperty CRC "2872004729"}
{attribute addProperty Size "9"}
TYPE SyncUnitTask_AB2F5079 EXTENDS SyncUnitTaskBase_FCD3CBF3 :
STRUCT
	{attribute addProperty Name "WcState"}
	WcState : WcState_0B2B16F9;
	{attribute addProperty Name "InfoData"}
	InfoData : InfoData_8649EEEB;
END_STRUCT
END_TYPE

// ---- Diagnostics/EtherCAT/SlaveDevice/Base/EtcSlaveBase_82538BE2.TcDUT

TYPE EtcSlaveBase_82538BE2 :
STRUCT
END_STRUCT
END_TYPE

// ---- Diagnostics/EtherCAT/SlaveDevice/Base/EtcSlaveBoxBase_77A0E4A7.TcDUT

{attribute clr[Container(Layout.Stack)]}
{attribute clr[Group(Layout.GroupBox)]}
{attribute addProperty PreviousPort "Unknown"}
{attribute addProperty SyncUnit "Unknown"}
TYPE EtcSlaveBoxBase_77A0E4A7 EXTENDS EtcSlaveBase_82538BE2 :
STRUCT
END_STRUCT
END_TYPE

// ---- Diagnostics/EtherCAT/SlaveDevice/Base/EtcSlaveEndTerminalBase_866C7F0C.TcDUT

{attribute clr[Container(Layout.Stack)]}
{attribute clr[Group(Layout.GroupBox)]}
{attribute addProperty PreviousPort "Unknown"}
{attribute addProperty SyncUnit "Unknown"}
TYPE EtcSlaveEndTerminalBase_866C7F0C EXTENDS EtcSlaveBase_82538BE2 :
STRUCT
END_STRUCT
END_TYPE

// ---- Diagnostics/EtherCAT/SlaveDevice/Base/EtcSlaveTerminalBase_947E5A46.TcDUT

{attribute clr[Container(Layout.Stack)]}
{attribute clr[Group(Layout.GroupBox)]}
{attribute addProperty PreviousPort "Unknown"}
{attribute addProperty SyncUnit "Unknown"}
TYPE EtcSlaveTerminalBase_947E5A46 EXTENDS EtcSlaveBase_82538BE2 :
STRUCT
END_STRUCT
END_TYPE

// ---- Diagnostics/EtherCAT/MasterDevice/InfoData_84133AC9.TcDUT
{attribute 'GeneratedUsingTerminal: IODEVICETYPE_ETHERCATPROT'}
{attribute addProperty BoxType "IODEVICETYPE_ETHERCATPROT"}
{attribute addProperty Id "ChangeCountAT %I*UINT2DevIdAT %I*UINT2AmsNetIdAT %I*AMSNETID6CfgSlaveCountAT %I*UINT2DcToTcTimeOffsetAT %I*LINT8DcToExtTimeOffsetAT %I*LINT8"}
{attribute addProperty CRC "3867959757"}
{attribute addProperty Size "28"}
TYPE InfoData_84133AC9 :
STRUCT
	{attribute addProperty Name "ChangeCount"}
	ChangeCount AT %I* : UINT;
	{attribute addProperty Name "DevId"}
	DevId AT %I* : UINT;
	{attribute addProperty Name "AmsNetId"}
	AmsNetId AT %I* : TcoAmsNetId;
	{attribute addProperty Name "CfgSlaveCount"}
	CfgSlaveCount AT %I* : UINT;
	{attribute addProperty Name "DcToTcTimeOffset"}
	DcToTcTimeOffset AT %I* : LINT;
	{attribute addProperty Name "DcToExtTimeOffset"}
	DcToExtTimeOffset AT %I* : LINT;
END_STRUCT
END_TYPE

// ---- Diagnostics/EtherCAT/MasterDevice/Inputs_A65FACA4.TcDUT
{attribute 'GeneratedUsingTerminal: IODEVICETYPE_ETHERCATPROT'}
{attribute addProperty BoxType "IODEVICETYPE_ETHERCATPROT"}
{attribute addProperty Id "SlaveCountAT %I*UINT2DevStateAT %I*UINT2Frm0StateAT %I*UINT2Frm0WcStateAT %I*UINT2Frm0InputToggleAT %I*UINT2"}
{attribute addProperty CRC "2791287972"}
{attribute addProperty Size "10"}
TYPE Inputs_A65FACA4 :
STRUCT
	{attribute addProperty Name "SlaveCount"}
	SlaveCount AT %I* : UINT;
	{attribute addProperty Name "DevState"}
	DevState AT %I* : UINT;
	{attribute addProperty Name "Frm0State"}
	Frm0State AT %I* : UINT;
	{attribute addProperty Name "Frm0WcState"}
	Frm0WcState AT %I* : UINT;
	{attribute addProperty Name "Frm0InputToggle"}
	Frm0InputToggle AT %I* : UINT;
END_STRUCT
END_TYPE

// ---- Diagnostics/EtherCAT/MasterDevice/Outputs_23C0ED1D.TcDUT
{attribute 'GeneratedUsingTerminal: IODEVICETYPE_ETHERCATPROT'}
{attribute addProperty BoxType "IODEVICETYPE_ETHERCATPROT"}
{attribute addProperty Id "DevCtrlAT %Q*UINT2Frm0CtrlAT %Q*UINT2Frm0WcCtrlAT %Q*UINT2"}
{attribute addProperty CRC "599846173"}
{attribute addProperty Size "6"}
TYPE Outputs_23C0ED1D :
STRUCT
	{attribute addProperty Name "DevCtrl"}
	DevCtrl AT %Q* : UINT;
	{attribute addProperty Name "Frm0Ctrl"}
	Frm0Ctrl AT %Q* : UINT;
	{attribute addProperty Name "Frm0WcCtrl"}
	Frm0WcCtrl AT %Q* : UINT;
END_STRUCT
END_TYPE

// ---- Diagnostics/EtherCAT/MasterDevice/TcoEthercatMasterDeviceState.TcDUT
TYPE TcoEthercatMasterDeviceState : STRUCT
	{attribute addProperty Name "Link error"}	
    LinkError : BOOL;
	{attribute addProperty Name "I/O locked after link error (I/O reset required)"}	
    IOLockedAfterLinkError : BOOL;
	{attribute addProperty Name "Link error (redundancy adapter)"}	
    LinkErrorRedundancyAdapter : BOOL;
	{attribute addProperty Name "Missing one frame (redundancy mode)"}	
    MissingOneFrame : BOOL;
	{attribute addProperty Name "Out of send resources (I/O reset required)"}	
    OutOfSendResources : BOOL;
	{attribute addProperty Name "Watchdog triggered"}	
    WatchdogTriggered : BOOL;
	{attribute addProperty Name "Ethernet driver (miniport) not found"}	
    EthernetDriverNotFound : BOOL;
	{attribute addProperty Name "I/O reset active"}	
    IOResetActive : BOOL;
	{attribute addProperty Name "At least one slave in 'INIT' state"}	
    AtLeastOneDeviceInInitState : BOOL;
	{attribute addProperty Name "At least one slave in 'PREOP' state"}	
    AtLeastOneDeviceInPreOpState : BOOL;
	{attribute addProperty Name "At least one slave in 'SAFEOP' state"}	
    AtLeastOneDeviceInSafeOpState : BOOL;
	{attribute addProperty Name "At least one device indicates an error state"}	
    AtLeastOneDeviceIndicatesAnErrorState : BOOL;
	{attribute addProperty Name "DC not in sync"}	
    DcNotInSync : BOOL;
END_STRUCT
END_TYPE

// ---- Diagnostics/EtherCAT/SlaveDevice/InfoData/InfoData_23CBA837.TcDUT
{attribute 'GeneratedUsingTerminal: EL6002-0000-0019'}
{attribute addProperty BoxType "EL6002-0000-0019"}
{attribute addProperty Id "AdsAddrAT %I*TcoIo.TcoAmsAddr0StateAT %I*UINT2"}
{attribute addProperty CRC "600549431"}
{attribute addProperty Size "2"}
TYPE InfoData_23CBA837 :
STRUCT
	{attribute addProperty Name "AdsAddr"}
	AdsAddr AT %I* : TcoAmsAddr;
	{attribute addProperty Name "State"}
	State AT %I* : UINT;
END_STRUCT
END_TYPE

// ---- Diagnostics/EtherCAT/SlaveDevice/InfoData/InfoData_6F19DB2B.TcDUT
{attribute 'GeneratedUsingTerminal: EL1809-0000-0018'}
{attribute addProperty BoxType "EL1809-0000-0018"}
{attribute addProperty Id "StateAT %I*UINT2"}
{attribute addProperty CRC "1863965483"}
{attribute addProperty Size "2"}
TYPE InfoData_6F19DB2B :
STRUCT
	{attribute addProperty Name "State"}
	State AT %I* : UINT;
END_STRUCT
END_TYPE

// ---- Diagnostics/EtherCAT/SlaveDevice/Inputs/InputBase_8311D824.TcDUT

TYPE InputBase_8311D824 :
STRUCT
END_STRUCT
END_TYPE

// ---- Diagnostics/EtherCAT/SlaveDevice/Outputs/OutputBase_10CEE7DE.TcDUT

TYPE OutputBase_10CEE7DE :
STRUCT
END_STRUCT
END_TYPE

// ---- Diagnostics/EtherCAT/SlaveDevice/WcState/WcState_0B2B16F9.TcDUT
{attribute 'GeneratedUsingTerminal: EL2809-0000-0018'}
{attribute addProperty BoxType "EL2809-0000-0018"}
{attribute addProperty Id "WcStateAT %I*BOOL1"}
{attribute addProperty CRC "187373305"}
{attribute addProperty Size "1"}
TYPE WcState_0B2B16F9 :
STRUCT
	{attribute addProperty Name "WcState"}
	WcState AT %I* : BOOL;
END_STRUCT
END_TYPE

// ---- Diagnostics/EtherCAT/SlaveDevice/WcState/WcState_9091E0EB.TcDUT
{attribute 'GeneratedUsingTerminal: EL6002-0000-0019'}
{attribute addProperty BoxType "EL6002-0000-0019"}
{attribute addProperty Id "WcStateAT %I*BOOL1InputToggleAT %I*BOOL1"}
{attribute addProperty CRC "2425479403"}
{attribute addProperty Size "2"}
TYPE WcState_9091E0EB :
STRUCT
	{attribute addProperty Name "WcState"}
	WcState AT %I* : BOOL;
	{attribute addProperty Name "InputToggle"}
	InputToggle AT %I* : BOOL;
END_STRUCT
END_TYPE

// ---- EtherCAT/eEcatState.TcDUT
{attribute 'qualified_only'}
TYPE eEcatState :
(
	MASK          := 15,
	INIT          := 1, 
	PREOP         := 2,  
	BOOTSTRAP     := 3,  
	SAFEOP        := 4,  
	OP            := 8,  
	ERROR         := 16,  
	INVALID_VPRS  := 32,  
	INITCMD_ERROR := 48,  
	DISABLED      := 128 
)BYTE;
END_TYPE

// ---- EtherCAT/eLinkState.TcDUT
{attribute 'qualified_only'}
TYPE eLinkState :
(
	EC_LINK_STATE_OK                := 0,
	EC_LINK_STATE_NOT_PRESENT       := 1,
	EC_LINK_STATE_LINK_WITHOUT_COMM := 2,
	EC_LINK_STATE_MISSING_LINK      := 4,
	EC_LINK_STATE_ADDITIONAL_LINK   := 8,
	EC_LINK_STATE_PORT_A            := 16,
	EC_LINK_STATE_PORT_B            := 32,
	EC_LINK_STATE_PORT_C            := 64,
	EC_LINK_STATE_PORT_D            := 128 			
)BYTE;
END_TYPE

// ---- SpecialPlcTypes/TcoAmsAddr.TcDUT
TYPE TcoAmsAddr :
	STRUCT
		netId : ARRAY [0..5] OF BYTE;
		port : WORD;
	END_STRUCT
END_TYPE

// ---- SpecialPlcTypes/TcoAmsNetId.TcDUT
TYPE TcoAmsNetId  :
	STRUCT
		netId : ARRAY [0..5] OF BYTE;
	END_STRUCT
END_TYPE

// ---- Diagnostics/EtherCAT/TcoEthercat.TcGVL
{attribute 'qualified_only'}
VAR_GLOBAL CONSTANT
    C_MaxSyncUnits : UINT := 10;
	C_MAX_LOCAL_ERROR_MESSAGES : UINT := 3;	
END_VAR

// ---- Diagnostics/EtherCAT/MasterDevice/SyncUnit/ITcoSyncUnit.TcIO
INTERFACE ITcoSyncUnit

PROPERTY DataInvalid : BOOL
GET
END_GET
END_PROPERTY

PROPERTY DataValid : BOOL
GET
END_GET
END_PROPERTY

PROPERTY HasSomeIssue : BOOL
GET
END_GET
END_PROPERTY

PROPERTY State : SyncUnitState
GET
END_GET
END_PROPERTY

END_INTERFACE

// ---- Diagnostics/EtherCAT/MasterDevice/ITcoEthercatMasterDevice.TcIO
INTERFACE ITcoEthercatMasterDevice

PROPERTY AllDataValid : BOOL
GET
END_GET
END_PROPERTY

PROPERTY DeviceHasSomeIssue : BOOL
GET
END_GET
END_PROPERTY

PROPERTY SomeDataInvalid : BOOL
GET
END_GET
END_PROPERTY

PROPERTY SomeSyncUnitHasSomeIssue : BOOL
GET
END_GET
END_PROPERTY

PROPERTY State : TcoEthercatMasterDeviceState
GET
END_GET
END_PROPERTY

END_INTERFACE

// ---- EtherCAT/ITcoEcatComponent.TcIO
INTERFACE ITcoEcatComponent

PROPERTY EcatState : REFERENCE TO TcoEcatSlaveState
GET
END_GET
END_PROPERTY

END_INTERFACE

// ---- POUs/MAIN.TcPOU
PROGRAM MAIN
VAR
END_VAR

END_PROGRAM

// ---- Diagnostics/EtherCAT/MasterDevice/SyncUnit/TcoSyncUnit.TcPOU
FUNCTION_BLOCK TcoSyncUnit EXTENDS TcoCore.TcoObject IMPLEMENTS ITcoSyncUnit
VAR
    {attribute addProperty Name "WcState"}
    WcState : WcState_0B2B16F9;
    {attribute addProperty Name "InfoData"}
    InfoData : InfoData_8649EEEB;
    {attribute addProperty Name "Status"}
    _State : SyncUnitState;
    {attribute 'hide'}
    _hasSomeIssue : BOOL;
    {attribute 'hide'}
    _dataValid : BOOL;
    {attribute 'hide'}
    _dataInvalid : BOOL;
END_VAR

PROPERTY DataInvalid : BOOL
GET
_dataInvalid := WcState.WcState;
DataInvalid := _dataInvalid;
END_GET
END_PROPERTY

PROPERTY DataValid : BOOL
GET
_dataValid := NOT WcState.WcState;
DataValid := _dataValid;
END_GET
END_PROPERTY

PROPERTY HasSomeIssue : BOOL
GET
VAR
	_syncUnitStatus : SyncUnitState;
END_VAR
_syncUnitStatus := State;

_hasSomeIssue := _syncUnitStatus.AtLeastOneSlaveInInitState OR
			_syncUnitStatus.AtLeastOneSlaveInPreopState OR
			_syncUnitStatus.AtLeastOneSlaveInBootState OR
			_syncUnitStatus.AtLeastOneSlaveInSafeOpState OR
			_syncUnitStatus.AtLeastOneSlaveSignalsError OR
			_syncUnitStatus.InvalidVendoridOrProductcodeRead OR
			_syncUnitStatus.InitializationErrorOccurred OR
			_syncUnitStatus.AtLeastOneSlaveNotPresent OR
			_syncUnitStatus.AtLeastOneSlaveSignalsLinkError OR
			_syncUnitStatus.AtLeastOneSlaveSignalsMissingLink OR
			_syncUnitStatus.AtLeastOneSlaveSignalsUnexpectedLink;
	
HasSomeIssue := _hasSomeIssue;
END_GET
END_PROPERTY

PROPERTY State : SyncUnitState
GET
_State.AtLeastOneSlaveInInitState := InfoData.State.0 AND NOT InfoData.State.1;
_State.AtLeastOneSlaveInPreopState := InfoData.State.0 AND InfoData.State.1;
_State.AtLeastOneSlaveInBootState := InfoData.State.0 AND InfoData.State.1;
_State.AtLeastOneSlaveInSafeOpState := InfoData.State.2;
_State.AtLeastOneSlaveInOpState := InfoData.State.3;
_State.AtLeastOneSlaveSignalsError := InfoData.State.4;
_State.InvalidVendoridOrProductcodeRead := InfoData.State.5;
_State.InitializationErrorOccurred := InfoData.State.6;
_State.AtLeastOneSlaveDisabled := InfoData.State.7;
_State.AtLeastOneSlaveNotPresent := InfoData.State.8;
_State.AtLeastOneSlaveSignalsLinkError := InfoData.State.9;
_State.AtLeastOneSlaveSignalsMissingLink := InfoData.State.10;
_State.AtLeastOneSlaveSignalsUnexpectedLink := InfoData.State.11;

State := _State;
END_GET
END_PROPERTY

END_FUNCTION_BLOCK

// ---- Diagnostics/EtherCAT/MasterDevice/Messenger/DiagnosticsMessenger.TcPOU
FUNCTION_BLOCK DiagnosticsMessenger EXTENDS TcoCore.TcoMessenger

{attribute 'hide'}
METHOD FB_init : BOOL
VAR_INPUT
	bInitRetains : BOOL; // if TRUE, the retain variables are initialized (warm start / cold start)
	bInCopyCode : BOOL;  // if TRUE, the instance afterwards gets moved into the copy code (online change)
	ParentObject : ITcoObject;
END_VAR
END_METHOD

END_FUNCTION_BLOCK

// ---- Diagnostics/EtherCAT/MasterDevice/Messenger/DiagnosticsMessengers.TcPOU
FUNCTION_BLOCK DiagnosticsMessengers EXTENDS TcoCore.TcoObject
VAR
	Messengers : ARRAY [0..2] OF DiagnosticsMessenger(THIS^);
END_VAR

{attribute 'hide'}
METHOD FB_init : BOOL
VAR_INPUT
	bInitRetains : BOOL; // if TRUE, the retain variables are initialized (warm start / cold start)
	bInCopyCode : BOOL;  // if TRUE, the instance afterwards gets moved into the copy code (online change)
	ParentObject : ITcoObject;	
END_VAR
Messengers[0].FB_init(bInitRetains,bInCopyCode,ParentObject);
Messengers[1].FB_init(bInitRetains,bInCopyCode,ParentObject);
Messengers[2].FB_init(bInitRetains,bInCopyCode,ParentObject);
END_METHOD

END_FUNCTION_BLOCK

// ---- Diagnostics/EtherCAT/MasterDevice/TcoEthercatDiagnosticsTask.TcPOU
FUNCTION_BLOCK TcoEthercatDiagnosticsTask EXTENDS TcoCore.TcoTask
VAR_INPUT
	inNetId : Tc2_System.T_AmsNetID;
END_VAR
VAR
    _EcGetAllSlaveStates 	: Tc2_EtherCAT.FB_EcGetAllSlaveStates;
    _EcGetConfSlaves 		: Tc2_EtherCAT.FB_EcGetConfSlaves;
	_updateDiagnosticsState : TcoCore.TcoState(THIS^,TcoCore.eRestoreMode.None);

	_SlaveStatesCount      		: UINT;
    _ConfigSlavesCount     		: UINT;
    _SlaveStateBuffer      		: ARRAY[0..EC_MAX_SLAVES] OF Tc2_EtherCAT.ST_EcSlaveState;
    _SlaveConfigDataBuffer 		: ARRAY[0..EC_MAX_SLAVES] OF Tc2_EtherCAT.ST_EcSlaveConfigData;

	_i	:	UINT;

	_name : STRING;
	_type : STRING;
	_state : STRING;
	
	_DiagnosticsMessengers		: DiagnosticsMessengers(THIS^);
	_DiagnosticsMessengerIndex	: UINT;	
END_VAR
VAR_OUTPUT
	outDiagnosticsAvailable : BOOL;
END_VAR

IF Execute() THEN
	IF _updateDiagnosticsState.State = 10 THEN
		outDiagnosticsAvailable := FALSE;
		_EcGetAllSlaveStates(bExecute := FALSE);
		_EcGetConfSlaves(bExecute := FALSE);
	
		IF NOT _EcGetAllSlaveStates.bBusy AND NOT _EcGetAllSlaveStates.bError AND NOT _EcGetConfSlaves.bBusy AND NOT _EcGetConfSlaves.bError THEN
			_updateDiagnosticsState.ChangeState(_updateDiagnosticsState._State + 10);
		END_IF
	END_IF
	
	IF _updateDiagnosticsState.State = 20 THEN
		_EcGetAllSlaveStates(sNetId := inNetId,
			pStateBuf := ADR(_SlaveStateBuffer),
			cbBufLen := SIZEOF(_SlaveStateBuffer),
			bExecute := TRUE,
			tTimeout :=,
			bBusy =>,
			bError =>,
			nErrId =>,
			nSlaves => _SlaveStatesCount);
	
		IF _EcGetAllSlaveStates.bBusy THEN
			_updateDiagnosticsState.ChangeState(_updateDiagnosticsState._State + 10);
		END_IF
	END_IF
	
	IF _updateDiagnosticsState.State = 30 THEN
		_EcGetAllSlaveStates(sNetId := inNetId,
			pStateBuf := ADR(_SlaveStateBuffer),
			cbBufLen := SIZEOF(_SlaveStateBuffer),
			bExecute := FALSE,
			tTimeout :=,
			bBusy =>,
			bError =>,
			nErrId =>,
			nSlaves => _SlaveStatesCount);
	
		IF NOT _EcGetAllSlaveStates.bBusy AND NOT _EcGetAllSlaveStates.bError THEN
			_updateDiagnosticsState.ChangeState(_updateDiagnosticsState._State + 10);
		END_IF
	END_IF
	
	IF _updateDiagnosticsState.State = 40 THEN
		_EcGetConfSlaves(sNetId := inNetId,
			pArrEcConfSlaveInfo := ADR(_SlaveConfigDataBuffer),
			cbBufLen := SIZEOF(_SlaveConfigDataBuffer),
			bExecute := TRUE,
			tTimeout :=,
			bBusy =>,
			bError =>,
			nErrorId =>,
			nSlaves => _ConfigSlavesCount);
	
		IF _EcGetConfSlaves.bBusy THEN
			_updateDiagnosticsState.ChangeState(_updateDiagnosticsState._State + 10);
		END_IF
	END_IF
	
	IF _updateDiagnosticsState.State = 50 THEN
		_EcGetConfSlaves(sNetId := inNetId,
			pArrEcConfSlaveInfo := ADR(_SlaveConfigDataBuffer),
			cbBufLen := SIZEOF(_SlaveConfigDataBuffer),
			bExecute := FALSE,
			tTimeout :=,
			bBusy =>,
			bError =>,
			nErrorId =>,
			nSlaves => _ConfigSlavesCount);
	
		IF NOT _EcGetConfSlaves.bBusy AND NOT _EcGetConfSlaves.bError THEN
			_updateDiagnosticsState.ChangeState(_updateDiagnosticsState._State + 10);
		END_IF
	END_IF
	
	IF _updateDiagnosticsState.State = 60 THEN
		_EcGetAllSlaveStates(bExecute := FALSE);
		_EcGetConfSlaves(bExecute := FALSE);
	
		IF NOT _EcGetAllSlaveStates.bBusy AND NOT _EcGetAllSlaveStates.bError AND NOT _EcGetConfSlaves.bBusy AND NOT _EcGetConfSlaves.bError THEN
			_updateDiagnosticsState.ChangeState(_updateDiagnosticsState._State + 10);
		END_IF
	END_IF
	
	IF _updateDiagnosticsState.State = 70 THEN
		_DiagnosticsMessengerIndex := 0;
	    FOR _i := 0 TO _ConfigSlavesCount DO
			IF (_SlaveStateBuffer[_i].deviceState <> 8 OR _SlaveStateBuffer[_i].linkState <> 0) THEN
				IF _SlaveConfigDataBuffer[_i].sName <> '' THEN
					IF _DiagnosticsMessengerIndex <= 2 THEN
						outDiagnosticsAvailable := TRUE;
						_name := _SlaveConfigDataBuffer[_i].sName;
						_type := Tc2_EtherCAT.F_ConvProductCodeToString(_SlaveConfigDataBuffer[_i].stSlaveIdentity);
						_state :=  Tc2_EtherCAT.F_ConvSlaveStateToString(state := _SlaveStateBuffer[_i]);
						_DiagnosticsMessengers.Messengers[_DiagnosticsMessengerIndex].Build().AppendAny(_name).Append('[').AppendAny(_type).Append(']').Append( _state).As().AsError().Pin();
						_DiagnosticsMessengerIndex := _DiagnosticsMessengerIndex + 1;
					END_IF
				END_IF
			END_IF;
	    END_FOR

		_updateDiagnosticsState.ChangeState(_updateDiagnosticsState._State + 10);
	END_IF
	
	IF _updateDiagnosticsState.State = 80 THEN
		DoneWhen(TRUE);
	END_IF

	ThrowWhen(_EcGetAllSlaveStates.bError OR _EcGetConfSlaves.bError);
END_IF

METHOD FB_init : BOOL
VAR_INPUT
	bInitRetains : BOOL; // if TRUE, the retain variables are initialized (warm start / cold start)
	bInCopyCode : BOOL;  // if TRUE, the instance afterwards gets moved into the copy code (online change)
	ParentObject : TcoCore.ITcoObject;	
END_VAR
END_METHOD

(*~
	<docu>
		<summary>
			Executes when task is aborted.
		</summary>			
	</docu>	
~*)
METHOD PROTECTED OnAbort
_EcGetAllSlaveStates(bExecute := FALSE);
_EcGetConfSlaves(bExecute := FALSE);

_updateDiagnosticsState.Restore();
END_METHOD

(*~
	<docu>
		<summary>
			Executes when task reaches the ```Done``` state .
		</summary>			
	</docu>	
~*)
METHOD PROTECTED OnDone
_EcGetAllSlaveStates(bExecute := FALSE);
_EcGetConfSlaves(bExecute := FALSE);
END_METHOD

(*~
	<docu>
		<summary>
			Executes when task reaches the ```Error``` state.
			<para>
				Do not confuse with <see cref="PlcDocu.TcoCore.TcoTask.WhileError()"/>, that is called cyclically until '''Error''' state is left.
			</para>
		</summary>			
	</docu>	
~*)
METHOD PROTECTED OnError
IF _EcGetAllSlaveStates.bError THEN
	Messenger.Build().Append('Reading status of all EtherCAT slaves using "Tc2_EtherCAT.FB_EcGetAllSlaveStates" function block returns error. nErrId: ').AppendAny(_EcGetAllSlaveStates.nErrId).As().AsError();
ELSIF _EcGetConfSlaves.bError THEN
	Messenger.Build().Append('Reading status of configurateed EtherCAT slaves using "Tc2_EtherCAT.FB_EcGetConfSlaves" function block returns error. nErrorId: ').AppendAny(_EcGetConfSlaves.nErrorId).As().AsError();
END_IF
END_METHOD

METHOD PROTECTED OnStart
_EcGetAllSlaveStates(bExecute := FALSE);
_EcGetConfSlaves(bExecute := FALSE);

_updateDiagnosticsState.ChangeState(10);
END_METHOD

(*~
	<docu>
		<summary>
			Restores this instance to the Ready state. Can be called explicitly or from within one of the restore mechanisms.
			<para>
				See also <see cref="PlcDocu.TcoCore.TcoTask.AutoRestorable()"/>
			</para>
		</summary>			
	</docu>	
~*)
METHOD Restore : ITcoRestorable
THIS^._EcGetAllSlaveStates(bExecute := FALSE);
THIS^._EcGetConfSlaves(bExecute := FALSE);

THIS^._DiagnosticsMessengers.Messengers[0].Clear();
THIS^._DiagnosticsMessengers.Messengers[1].Clear();
THIS^._DiagnosticsMessengers.Messengers[2].Clear();

THIS^.outDiagnosticsAvailable := FALSE;
THIS^._updateDiagnosticsState.Restore();

SUPER^.Restore();
END_METHOD

END_FUNCTION_BLOCK

// ---- Diagnostics/EtherCAT/MasterDevice/TcoEthercatMasterDevice.TcPOU
FUNCTION_BLOCK TcoEthercatMasterDevice EXTENDS TcoCore.TcoComponent IMPLEMENTS ITcoEthercatMasterDevice
VAR_INPUT
    Inputs   		:	Inputs_A65FACA4;
    InfoData		:	InfoData_84133AC9;
	SyncUnits		:	POINTER TO SyncUnitTask_AB2F5079;
	SyncUnitsSize	:	UINT;
END_VAR

VAR
    _someSyncUnitHasSomeIssue	: BOOL;
    _allDataValid          		: BOOL;
    _someDataInvalid       		: BOOL;
    _State                		: TcoEthercatMasterDeviceState;
    _NetId                 		: Tc2_System.T_AmsNetID;
    _DeviceHasSomeIssue    		: BOOL;
    _TcoEthercatDiagnosticsTask	: TcoEthercatDiagnosticsTask(THIS^);

    _InfoDataChangeCountPV 		: UINT;

	_numberOfSyncUnits			: UINT;

	{attribute addProperty Name "Acknowledge"}
	_acknowledge				:	TcoCore.TcoTask(THIS^);
	
	_DiagnosticsAvailable : BOOL;
END_VAR
VAR_OUTPUT
    Outputs  : Outputs_23C0ED1D;
END_VAR

UpdateSyncUnitsStatus(SyncUnits,SyncUnitsSize);
Diagnostics();

PROPERTY AllDataValid : BOOL
GET
AllDataValid := _allDataValid;
END_GET
END_PROPERTY

PROPERTY DeviceHasSomeIssue : BOOL
GET
_DeviceHasSomeIssue		:=	_State.LinkError							 	OR
							_State.IOLockedAfterLinkError 					OR
							_State.LinkErrorRedundancyAdapter	 			OR
							_State.MissingOneFrame 							OR
							_State.OutOfSendResources 						OR
							_State.WatchdogTriggered 						OR
							_State.EthernetDriverNotFound 					OR
							_State.IOResetActive 							OR
							_State.AtLeastOneDeviceInInitState 				OR
							_State.AtLeastOneDeviceInPreOpState 			OR
							_State.AtLeastOneDeviceInSafeOpState 			OR
							_State.AtLeastOneDeviceIndicatesAnErrorState 	OR
							_State.DcNotInSync 								;
							
DeviceHasSomeIssue := _DeviceHasSomeIssue;
END_GET
END_PROPERTY

METHOD Diagnostics
VAR
    _i : UINT;
END_VAR
_NetId := Tc2_System.F_CreateAmsNetId(InfoData.AmsNetId.netId);

_TcoEthercatDiagnosticsTask(inNetId := _NetId, outDiagnosticsAvailable => _DiagnosticsAvailable);

Service();

IF _acknowledge.Execute() THEN
	Restore();	
END_IF

IF (DeviceHasSomeIssue OR SomeSyncUnitHasSomeIssue OR SomeDataInvalid OR _InfoDataChangeCountPV <> InfoData.ChangeCount) (*OR _manualDiagnosticStart.Execute()*) THEN
	IF _TcoEthercatDiagnosticsTask.Ready THEN
		_InfoDataChangeCountPV := InfoData.ChangeCount;
		_TcoEthercatDiagnosticsTask.Invoke();
	END_IF
	IF _TcoEthercatDiagnosticsTask.Done AND NOT _DiagnosticsAvailable THEN
		_TcoEthercatDiagnosticsTask.Restore();
	END_IF;
END_IF
END_METHOD

METHOD FB_init : BOOL
VAR_INPUT
	bInitRetains : BOOL; // if TRUE, the retain variables are initialized (warm start / cold start)
	bInCopyCode : BOOL;  // if TRUE, the instance afterwards gets moved into the copy code (online change)
	ParentObject : TcoCore.ITcoObject;	
END_VAR
END_METHOD

(*~
	<docu>
		<summary>
			Restores this instance to the Ready state. Can be called explicitly or from within one of the restore mechanisms.	
		</summary>			
	</docu>	
~*)
METHOD  Restore : ITcoRestorable
THIS^.Messenger.Clear();
THIS^._DiagnosticsAvailable := FALSE;
THIS^._acknowledge.Restore();
THIS^._TcoEthercatDiagnosticsTask.Restore();
END_METHOD

(*~
	<docu>
		<summary>
		    Custom service (manual, maintenance) logic.
			This method must be implemented in derived class.
		</summary>			
	</docu>	
~*)
METHOD PROTECTED  ServiceMode
_acknowledge();
END_METHOD

PROPERTY SomeDataInvalid : BOOL
GET
SomeDataInvalid := _someDataInvalid;
END_GET
END_PROPERTY

PROPERTY SomeSyncUnitHasSomeIssue : BOOL
GET
SomeSyncUnitHasSomeIssue := _someSyncUnitHasSomeIssue;
END_GET
END_PROPERTY

PROPERTY State : TcoEthercatMasterDeviceState
GET
_State.LinkError							 	:= Inputs.DevState.0;
_State.IOLockedAfterLinkError 					:= Inputs.DevState.1;
_State.LinkErrorRedundancyAdapter	 			:= Inputs.DevState.2;
_State.MissingOneFrame 							:= Inputs.DevState.3;
_State.OutOfSendResources 						:= Inputs.DevState.4;
_State.WatchdogTriggered 						:= Inputs.DevState.5;
_State.EthernetDriverNotFound 					:= Inputs.DevState.6;
_State.IOResetActive 							:= Inputs.DevState.7;
_State.AtLeastOneDeviceInInitState 				:= Inputs.DevState.8;
_State.AtLeastOneDeviceInPreOpState 			:= Inputs.DevState.9;
_State.AtLeastOneDeviceInSafeOpState 			:= Inputs.DevState.10;
_State.AtLeastOneDeviceIndicatesAnErrorState 	:= Inputs.DevState.11;
_State.DcNotInSync 								:= Inputs.DevState.12;

State := _State;
END_GET
END_PROPERTY

METHOD SyncUnitHasSomeIssue : BOOL
VAR_INPUT
	inState : UINT;
END_VAR
VAR
	_state : SyncUnitState;
END_VAR
_state.AtLeastOneSlaveInInitState 				:=	inState.0 AND NOT	inState.1;
_state.AtLeastOneSlaveInPreopState 				:=	inState.0 AND 		inState.1;
_state.AtLeastOneSlaveInBootState 				:=	inState.0 AND		inState.1;
_state.AtLeastOneSlaveInSafeOpState 			:=	inState.2;
_state.AtLeastOneSlaveInOpState 				:=	inState.3;
_state.AtLeastOneSlaveSignalsError 				:=	inState.4;
_state.InvalidVendoridOrProductcodeRead 		:=	inState.5;
_state.InitializationErrorOccurred				:=	inState.6;
_state.AtLeastOneSlaveDisabled					:=	inState.7;
_state.AtLeastOneSlaveNotPresent				:=	inState.8;
_state.AtLeastOneSlaveSignalsLinkError			:=	inState.9;
_state.AtLeastOneSlaveSignalsMissingLink		:=	inState.10;
_state.AtLeastOneSlaveSignalsUnexpectedLink		:=	inState.11;

SyncUnitHasSomeIssue :=	_state.AtLeastOneSlaveInInitState OR
						_state.AtLeastOneSlaveInPreopState OR
						_state.AtLeastOneSlaveInBootState OR
						_state.AtLeastOneSlaveInSafeOpState OR
						_state.AtLeastOneSlaveSignalsError OR
						_state.InvalidVendoridOrProductcodeRead OR
						_state.InitializationErrorOccurred OR
						_state.AtLeastOneSlaveNotPresent OR
						_state.AtLeastOneSlaveSignalsLinkError OR
						_state.AtLeastOneSlaveSignalsMissingLink OR
						_state.AtLeastOneSlaveSignalsUnexpectedLink;
END_METHOD

METHOD UpdateSyncUnitsStatus
VAR_INPUT
	SyncUnits			:	POINTER TO SyncUnitTask_AB2F5079;
	SyncUnitsSize		:	UINT;
END_VAR
VAR
    _i					:	UINT;
	_pSyncUnit			:	POINTER TO SyncUnitTask_AB2F5079;
	_SyncUnit			:	SyncUnitTask_AB2F5079;
	_SyncUnitState		:	UINT;
END_VAR
_someSyncUnitHasSomeIssue := FALSE;
_allDataValid := TRUE;
_someDataInvalid := FALSE;

IF SyncUnits<>0 THEN
	_numberOfSyncUnits := SyncUnitsSize / SIZEOF(SyncUnitTask_AB2F5079);
	FOR _i := 0 TO _numberOfSyncUnits - 1 DO
		_pSyncUnit					:=	SyncUnits + _i * SIZEOF(SyncUnitTask_AB2F5079);
		_SyncUnit					:=	_pSyncUnit^;	
		_someSyncUnitHasSomeIssue 	:=	_someSyncUnitHasSomeIssue OR SyncUnitHasSomeIssue(_SyncUnit.InfoData.State);
		_allDataValid				:=	_allDataValid AND NOT _SyncUnit.WcState.WcState;
		_someDataInvalid			:=	_someDataInvalid OR _SyncUnit.WcState.WcState;
	END_FOR
END_IF
END_METHOD

END_FUNCTION_BLOCK

// ---- Diagnostics/ProfinetComponent/TcoPnIoComponent.TcPOU
FUNCTION_BLOCK ABSTRACT TcoPnIoComponent EXTENDS TcoCore.TcoComponent
VAR_INPUT
	inPnIoBoxState : UINT;
	inPnIoBoxDiag : UINT;
END_VAR
VAR
	 //*{attribute addProperty Name "<#PN ready#>"}
     //*{attribute clr [ReadOnly()]}
	_profinetReady : BOOL;
END_VAR

//PnIoBoxState
//0 = No error
//1 = Profinet device state machine is in boot mode
//2 = Device not found
//3 = The stationname is not unique
//4 = IP could not be set
//5 = IP conflict
//6 = DCP set was not successful
//7 = Watchdog error
//8 = Datahold error
//9 = RTC3: Sync mode could not be initiated
//10 = Profinet controller has a link error
//11 = The aliasname is not unique
//12 = The automatic name assignement isn't possible - wrong device type
//13 = IOC-AR is established but no application ready
//14 = IOC-AR is established but module difference
//15 = At least one InputCR is invalid, provider in stop or problemindicator is set
//16 = At least one OutputCR is invalid, provider in stop or problemindicator is set
//31 = Only for EtherCAT gateways: WC-State of cyclic EtherCAT frame is 1

THIS^.Messenger.OnCondition(inPnIoBoxState=1 ).Error('<#Profinet device state machine is in boot mode!#>'); 
THIS^.Messenger.OnCondition(inPnIoBoxState=2 ).Error('<#Device NOT found!#>'); 
THIS^.Messenger.OnCondition(inPnIoBoxState=3 ).Error('<#The stationname is not unique!#>'); 
THIS^.Messenger.OnCondition(inPnIoBoxState=4 ).Error('<#IP could NOT be set!#>'); 
THIS^.Messenger.OnCondition(inPnIoBoxState=5 ).Error('<#IP conflict!#>'); 
THIS^.Messenger.OnCondition(inPnIoBoxState=6 ).Error('<#DCP set was NOT successful!#>'); 
THIS^.Messenger.OnCondition(inPnIoBoxState=7 ).Error('<#Watchdog error!#>'); 
THIS^.Messenger.OnCondition(inPnIoBoxState=8 ).Error('<#Datahold error!#>'); 
THIS^.Messenger.OnCondition(inPnIoBoxState=9 ).Error('<#RTC3: Sync mode could not be initiated!#>'); 
THIS^.Messenger.OnCondition(inPnIoBoxState=10).Error('<#Profinet controller has a link error!#>'); 
THIS^.Messenger.OnCondition(inPnIoBoxState=11).Error('<#The aliasname is not unique!#>'); 
THIS^.Messenger.OnCondition(inPnIoBoxState=12).Error('<#The automatic name assignement is not possible - wrong device TYPE!#>'); 
THIS^.Messenger.OnCondition(inPnIoBoxState=13).Error('<#IOC-AR is established but no application ready!#>'); 
THIS^.Messenger.OnCondition(inPnIoBoxState=14).Error('<#IOC-AR is established but module difference!#>'); 
THIS^.Messenger.OnCondition(inPnIoBoxState=15).Error('<#AT least one InputCR is invalid, provider in stop OR problemindicator is set!#>'); 
THIS^.Messenger.OnCondition(inPnIoBoxState=16).Error('<#At least one OutputCR is invalid, provider in stop or problemindicator is set!#>'); 
THIS^.Messenger.OnCondition(inPnIoBoxState=31).Error('<#EtherCAT gateway: WC-State OF cyclic EtherCAT frame is 1!#>'); 

//PnIoBoxDiag
//0x0000 = No diagnosis
//0x0001 = IOC-AR is not established
//0x0002 = IOC-AR is established
//0x0004 = IOC-AR is established but no application ready
//0x0008 = IOC-AR is established but module difference
//0x0010 = At least one AlarmCR got a diagnosis alarm
//0x0100 = At least one InputCR is invalid
//0x0200 = At least one InputCR Provider is in stop
//0x0400 = At least one InputCR Problemindicator is set
//0x1000 = At least one OutputCR is invalid
//0x2000 = At least one OutputCR Provider is in stop
//0x4000 = At least one OutputCR Problemindicator is set

THIS^.Messenger.OnCondition(inPnIoBoxDiag.0 ).Error('<#IOC-AR is not established!#>'); 
THIS^.Messenger.OnCondition(NOT _profinetReady AND inPnIoBoxDiag.1 ).Info('<#IOC-AR is established!#>');
THIS^.Messenger.OnCondition(inPnIoBoxDiag.2 ).Error('<#IOC-AR is established but no application ready!#>');
THIS^.Messenger.OnCondition(inPnIoBoxDiag.3 ).Error('<#IOC-AR is established but module difference!#>');
THIS^.Messenger.OnCondition(inPnIoBoxDiag.4 ).Error('<#AT least one AlarmCR got a diagnosis alarm!#>');
THIS^.Messenger.OnCondition(inPnIoBoxDiag.8 ).Error('<#At least one InputCR is invalid!#>');
THIS^.Messenger.OnCondition(inPnIoBoxDiag.9 ).Error('<#AT least one InputCR Provider is in stop!#>');
THIS^.Messenger.OnCondition(inPnIoBoxDiag.10).Error('<#At least one InputCR Problemindicator is set!#>');
THIS^.Messenger.OnCondition(inPnIoBoxDiag.12).Error('<#AT least one OutputCR is invalid!#>');
THIS^.Messenger.OnCondition(inPnIoBoxDiag.13).Error('<#At least one OutputCR Provider is in stop!#>');
THIS^.Messenger.OnCondition(inPnIoBoxDiag.14).Error('<#AT least one OutputCR Problemindicator is set!#>');


_profinetReady := inPnIoBoxState = 0 AND inPnIoBoxDiag = 2;

PROPERTY ProfinetReady : BOOL
GET
ProfinetReady := _profinetReady;
END_GET
END_PROPERTY

END_FUNCTION_BLOCK

// ---- EtherCAT/TcoEcatSlaveState.TcPOU
FUNCTION_BLOCK  TcoEcatSlaveState EXTENDS TcoObject 
VAR_INPUT
    AdsAddr : AMSADDR;
END_VAR
VAR_OUTPUT
END_VAR
VAR

    //*	{attribute addProperty Name "<#Actual state#>"}
    //*	{attribute clr [ReadOnly()]}
    _ecatState : eEcatState;
    //*	{attribute addProperty Name "<#Actual Link state#>"}
    //*	{attribute clr [ReadOnly()]}
    _linkState : eLinkState;
    //*	{attribute addProperty Name "<#ECAT Communication Ok#>"}
    //*	{attribute clr [ReadOnly()]}
    _ecatOk : BOOL;
 
    //*	{attribute clr [RenderIgnore()]}
    _progress : INT := 0;
	

    //*	{attribute addProperty Name "<#EtherCat masters Ams Net Id#>"}
    //*	{attribute clr [ReadOnly()]}
    _netId : STRING[23]; //as string	

	 //* {attribute clr [RenderIgnore()]}
    _etherCAT_Addr : UINT;

	//*	{attribute addProperty Name "<#State check Time(Period)#>"}
   	_periodStateCheckTime: TIME :=T#1S;
	
	//*	{attribute addProperty Name "<#Error Time#>"}
   	_errorTime: TIME :=T#5S;
    //*	{attribute clr [RenderIgnore()]}
    _getSlaveState : FB_EcGetSlaveState;
    //*	{attribute clr [RenderIgnore()]}
    _setSlaveState : FB_EcSetSlaveState;


    //*	{attribute clr [RenderIgnore()]}
    bExecute : BOOL;
    //*	{attribute clr [RenderIgnore()]}
    state : ST_EcSlaveState;
    //*	{attribute clr [RenderIgnore()]}
    _error : BOOL;
    //*	{attribute clr [RenderIgnore()]}
    _busy : BOOL;
    //*	{attribute clr [RenderIgnore()]}
    _errId : UDINT;
    //*	{attribute clr [RenderIgnore()]}
    _stateTimer : TON;
	//*	{attribute clr [RenderIgnore()]}
    _errorTimer : TON;
	
    //*	{attribute addProperty Name "<#Required state#>"}
    _ecatReqestState : eEcatState;
	
    //*	{attribute addProperty Name "<#Change State#>"}
    _changeStateTask : TcoCore.TcoTask(THIS^);

    //*	{attribute addProperty Name "<#Restore#>"}
    _restoreTask : TcoCore.TcoTask(THIS^);

	 {attribute 'hide'} 
	_sb : TcoCore.StringBuilder;
	{attribute 'hide'} 
	_amsEmpty: BOOL;
END_VAR

_netId := F_CreateAmsNetId(nIds := AdsAddr.netId);
_etherCAT_Addr := AdsAddr.port;
_amsEmpty:=(_netId = '0.0.0.0.0.0') OR (_etherCAT_Addr = 0);
	

IF _changeStateTask.Execute() THEN
	_changeStateTask.DoneWhen(ChangeState(RequestedDeviceState:=_ecatReqestState ));
END_IF

THIS^._changeStateTask.ThrowWhen((_changeStateTask.ElapsedTime>=_errorTime AND _progress>0) 
								OR _amsEmpty ); 

THIS^._changeStateTask.Messenger.OnCondition(_amsEmpty).Error('<#Ads address information is not defined!#>');
//*************RESTORE********************

_restoreTask.Enabled := TRUE;
IF _restoreTask.Execute() THEN
	Restore();
END_IF
//****************************************


IF (_amsEmpty) THEN		
	RETURN;
END_IF


THIS^._GetState(_periodStateCheckTime);

METHOD PRIVATE _GetState
VAR_INPUT
	Period:TIME;
END_VAR
_stateTimer(IN := TRUE,PT := Period);		

IF _stateTimer.Q THEN
	bExecute := TRUE;
	_stateTimer(IN := FALSE);
END_IF
 
_getSlaveState(sNetId:= _netId, 
				nSlaveAddr := _etherCAT_Addr, 
				bExecute := bExecute,
				bBusy => _busy,
				state => state,
				bError => _error,
				nErrId => _ErrId);

IF NOT _busy THEN
	_ecatState := state.deviceState;
	_linkState := state.linkState;
	_ecatOk := (state.deviceState = EC_DEVICE_STATE_OP);
	bExecute := FALSE;
END_IF
END_METHOD

PROPERTY PUBLIC EcatOk : BOOL
GET
EcatOk:=_ecatOk;
END_GET
END_PROPERTY

PROPERTY PUBLIC ErrorTime : TIME
GET
ErrorTime:=_errorTime;
END_GET
SET
_errorTime:=ErrorTime;
END_SET
END_PROPERTY

METHOD PUBLIC ChangeState : BOOL
VAR_INPUT
	RequestedDeviceState:BYTE;
END_VAR
ChangeState := FALSE;

_setSlaveState(sNetId := _netId,
    nSlaveAddr := _etherCAT_Addr,
    bExecute :=,
    tTimeout :=,
    reqState :=,
    bBusy =>,
    bError =>,
    nErrId =>,
    currState => state);

CASE _progress OF
    0:
        _ecatOk := FALSE;
        _setSlaveState(bExecute := FALSE);
        _progress := 10;

    10:
        _setSlaveState(reqState := EC_DEVICE_STATE_INIT);
        _setSlaveState(bExecute := TRUE);

        IF _setSlaveState.bBusy THEN
            _progress := 15;
        END_IF
    15: //INIT
        IF (state.deviceState) = EC_DEVICE_STATE_INIT AND
            RequestedDeviceState > state.deviceState AND
            RequestedDeviceState <> EC_DEVICE_STATE_BOOTSTRAP THEN
            _setSlaveState(bExecute := FALSE);
            _progress := 30;
        ELSIF (state.deviceState) = EC_DEVICE_STATE_INIT AND
            RequestedDeviceState > state.deviceState AND
            RequestedDeviceState = EC_DEVICE_STATE_BOOTSTRAP THEN
            _setSlaveState(bExecute := FALSE);
            _progress := 20;
        ELSIF NOT _setSlaveState.bBusy AND (state.deviceState) = RequestedDeviceState THEN
            _progress := 100;

        END_IF

    20:
        _setSlaveState(reqState := EC_DEVICE_STATE_BOOTSTRAP);
        _setSlaveState(bExecute := TRUE);

        IF _setSlaveState.bBusy THEN
            _progress := 25;
        END_IF
    25: ///BOOTSTRAP
        IF (state.deviceState) = EC_DEVICE_STATE_BOOTSTRAP THEN
            _setSlaveState(bExecute := FALSE);
            _progress := 100;
        END_IF

    30:
        _setSlaveState(reqState := EC_DEVICE_STATE_PREOP);
        _setSlaveState(bExecute := TRUE);

        IF _setSlaveState.bBusy THEN
            _progress := 35;
        END_IF
    35: //PREOP
        IF (state.deviceState) = EC_DEVICE_STATE_PREOP AND RequestedDeviceState > state.deviceState THEN
            _setSlaveState(bExecute := FALSE);
            _progress := 40;
        ELSIF NOT _setSlaveState.bBusy AND (state.deviceState) = RequestedDeviceState THEN
            _progress := 100;
        END_IF

    40:
        _setSlaveState(reqState := EC_DEVICE_STATE_SAFEOP);
        _setSlaveState(bExecute := TRUE);

        IF _setSlaveState.bBusy THEN
            _progress := 45;
        END_IF
    45: //SAFEOP
        IF (state.deviceState) = EC_DEVICE_STATE_SAFEOP AND RequestedDeviceState > state.deviceState THEN
            _setSlaveState(bExecute := FALSE);
            _progress := 50;
        ELSIF NOT _setSlaveState.bBusy AND (state.deviceState) = RequestedDeviceState THEN
            _progress := 100;
        END_IF

    50: //OP
        _setSlaveState(reqState := EC_DEVICE_STATE_OP);
        _setSlaveState(bExecute := TRUE);

        IF (state.deviceState) = EC_DEVICE_STATE_OP THEN
            _setSlaveState(bExecute := FALSE);
            _ecatOk := TRUE;
            _progress := 100;

        END_IF

    100:

        ChangeState := TRUE;
        _progress := 0;

END_CASE
Messenger.OnCondition(NOT _setSlaveState.bBusy AND RequestedDeviceState > EC_DEVICE_STATE_OP)
    .Post(_sb.Clear().Append('<#Unexpected state: #>').Append(TO_STRING(state.deviceState)).ToString(), eMessageCategory.Error);
END_METHOD

PROPERTY PUBLIC ChangeStateTask : TcoCore.ITcoTaskStatus
GET
ChangeStateTask:=_changeStateTask;
END_GET
END_PROPERTY

PROPERTY PUBLIC PeriodCheckState : TIME
GET
PeriodCheckState:= _periodStateCheckTime;
END_GET
SET
_periodStateCheckTime:=PeriodCheckState;
END_SET
END_PROPERTY

METHOD Restore  : ITcoRestorable
VAR_INPUT
END_VAR
_changeStateTask.Restore();
_ecatOk:=false;
_progress:=0;
_restoreTask.Restore();
END_METHOD

END_FUNCTION_BLOCK

// ---- EtherCAT/TcoEcatComponent.TcPOU
FUNCTION_BLOCK ABSTRACT TcoEcatComponent EXTENDS TcoCore.TcoComponent IMPLEMENTS ITcoEcatComponent
VAR_INPUT
    AdsAddr : AMSADDR;
END_VAR
VAR_OUTPUT
END_VAR
VAR
	//*	{attribute addProperty Name "<#Ecat slave state#>"}
	_ecatState:TcoEcatSlaveState(THIS^);
	{attribute 'hide'} 
	_sb : TcoCore.StringBuilder;

END_VAR

_ecatState(AdsAddr:=AdsAddr);

PROPERTY PUBLIC EcatState : REFERENCE TO TcoEcatSlaveState
GET
EcatState REF=_ecatState;
END_GET
END_PROPERTY

METHOD Restore  : ITcoRestorable
VAR_INPUT
END_VAR
_ecatState.Restore();
END_METHOD

METHOD PROTECTED  ServiceMode
VAR_INPUT
END_VAR
END_METHOD

END_FUNCTION_BLOCK
